END_VAR
VAR CONSTANT
	unWaitInterrupt						:UINT := 0;
	unDuringInterrupt						:UINT := 1;
	unAfterInterrupt						:UINT := 2;
	unChkFile							:UINT := 3;
	unNoInterrupt							:UINT := 4;
END_VAR

IF NOT bEnable
THEN
	bBusy := FALSE;
	bDone := FALSE;
	bError := FALSE;
	bEStop := FALSE;
	bFirstTime := FALSE;
	RETURN;
END_IF

IF NOT bFirstTime
THEN
	bBusy := FALSE;
	bDone := FALSE;
	bError := FALSE;
	bEStop := FALSE;
	unState := 0;
	unIncLog := 1;
	unIncDuringInterrupt := 1;
	unIncAfterInterrupt := 1;

	unLOG_INSTANCE_IDX  := GVL_Logger.unLOG_INSTANCE_IDX + 1;
	unInstanceIdx := unLOG_INSTANCE_IDX;

	unState := unWaitInterrupt;

	bFirstTime := TRUE;
END_IF


rtDeleteAll(CLK := bDeleteAll);

IF rtDeleteAll.Q
    AND (bDone OR bError)
THEN
	bBusy := FALSE;
	bDone := FALSE;
	bError := FALSE;
	bEStop := FALSE;
	unState := 0;
	unIncLog := 1;
	unIncDuringInterrupt := 1;
	unIncAfterInterrupt := 1;

	unState := unWaitInterrupt;
END_IF

rtInterrupt(CLK := bInterrupt);
IF rtInterrupt.Q
THEN
	unState := unWaitInterrupt;
END_IF;

udnCycleNo := udnCycleNo + 1;

CASE unState OF
	
	unWaitInterrupt:
		bBusy := FALSE;
		bDone := FALSE;
		bError := FALSE;

		fbLoggerFile.bExecute := FALSE;

		(* Shift down logger list by 1 *)
		A_ShiftDown();

		(* Write time stamp and value of variables before interrupt *)
		arstLoggerWaitInterrupt[1].udnCycleNo := udnCycleNo;
		arstLoggerWaitInterrupt[1].sTimeStamp := sDateTime;
		arstLoggerWaitInterrupt[1].arsLogVars := arsLogVars;

		IF bInterrupt
		THEN
			bBusy := TRUE;
			bDone := FALSE;

			bEStop := bLogOne;

			MEMSET(ADR(arstLoggerDuringInterrupt), 0, SIZEOF(arstLoggerDuringInterrupt));
			MEMSET(ADR(arstLoggerAfterInterrupt), 0, SIZEOF(arstLoggerAfterInterrupt));

			(* Log data *)
			IF unIncLog <= GVL_Logger.unLOG_MAX_NO
			THEN
				MEMCPY(ADR(arstLogger[unIncLog].arstLoggerWaitInterrupt), ADR(arstLoggerWaitInterrupt), SIZEOF(arstLoggerWaitInterrupt));
			ELSE
				unIncLog := 1;
				MEMCPY(ADR(arstLogger[unIncLog].arstLoggerWaitInterrupt), ADR(arstLoggerWaitInterrupt), SIZEOF(arstLoggerWaitInterrupt));
			END_IF

			(* Write time stamp and value of variables during interrupt *)
			unIncDuringInterrupt := 1;
			arstLoggerDuringInterrupt[unIncDuringInterrupt].udnCycleNo := udnCycleNo;
			arstLoggerDuringInterrupt[unIncDuringInterrupt].sTimeStamp := sDateTime;
			arstLoggerDuringInterrupt[unIncDuringInterrupt].arsLogVars := arsLogVars;
			unIncDuringInterrupt := unIncDuringInterrupt + 1;

			fbLoggerFile.sFileName := CONCAT(
										sDateTime,
										CONCAT(
											'_',
											UINT_TO_STRING(unInstanceIdx)
										)
									);

			unState := unDuringInterrupt;

		END_IF

	unDuringInterrupt:
		IF unIncDuringInterrupt <= GVL_Logger.unLOG_DURING_MAX_NO
		THEN
			(*  Write time stamp and value of variables during interrupt *)
			arstLoggerDuringInterrupt[unIncDuringInterrupt].udnCycleNo := udnCycleNo;
			arstLoggerDuringInterrupt[unIncDuringInterrupt].sTimeStamp := sDateTime;
			arstLoggerDuringInterrupt[unIncDuringInterrupt].arsLogVars := arsLogVars;
		
			unIncDuringInterrupt := unIncDuringInterrupt + 1;

		END_IF

		IF NOT bInterrupt
		THEN
			(* Log data *)
			MEMCPY(ADR(arstLogger[unIncLog].arstLoggerDuringInterrupt), ADR(arstLoggerDuringInterrupt), SIZEOF(arstLoggerDuringInterrupt));

			(* Write time stamp and value of variables after interrupt *)
			unIncAfterInterrupt := 1;
			arstLoggerAfterInterrupt[unIncAfterInterrupt].udnCycleNo := udnCycleNo;
			arstLoggerAfterInterrupt[unIncAfterInterrupt].sTimeStamp := sDateTime;
			arstLoggerAfterInterrupt[unIncAfterInterrupt].arsLogVars := arsLogVars;
			unIncAfterInterrupt := unIncAfterInterrupt + 1;

			unState := unAfterInterrupt;

		END_IF

	unAfterInterrupt:
		IF unIncAfterInterrupt <= GVL_Logger.unLOG_AFTER_MAX_NO
		THEN
			(* Write time stamp and value of variables after interrupt *)
			arstLoggerAfterInterrupt[unIncAfterInterrupt].udnCycleNo := udnCycleNo;
			arstLoggerAfterInterrupt[unIncAfterInterrupt].sTimeStamp := sDateTime;	
			arstLoggerAfterInterrupt[unIncAfterInterrupt].arsLogVars := arsLogVars;

			unIncAfterInterrupt := unIncAfterInterrupt + 1;
		ELSE
			(* Log data *)
			MEMCPY(ADR(arstLogger[unIncLog].arstLoggerAfterInterrupt), ADR(arstLoggerAfterInterrupt), SIZEOF(arstLoggerAfterInterrupt));

			fbLoggerFile.bExecute := TRUE;

			IF fbLoggerFile.bBusy
			THEN
				unState := unChkFile;

			ELSIF fbLoggerFile.bError
			THEN
				fbLoggerFile.bExecute := FALSE;
	
				bBusy := FALSE;
				bError := TRUE;
	
				unState := unNoInterrupt;

			END_IF
		END_IF

	unChkFile:
		IF NOT bEnableSaveInFile
		     OR fbLoggerFile.bDone
		THEN
			fbLoggerFile.bExecute := FALSE;

			bBusy := FALSE;
			bDone := TRUE;

			unState := unNoInterrupt;

		ELSIF  fbLoggerFile.bError
		THEN
			fbLoggerFile.bExecute := FALSE;

			bBusy := FALSE;
			bError := TRUE;

			unState := unNoInterrupt;

		END_IF

	unNoInterrupt:
		IF NOT bInterrupt
		    AND NOT bEStop
		THEN
			bBusy := FALSE;
			bDone := FALSE;
			bError := FALSE;

			unIncLog := unIncLog + 1;

			unState := unWaitInterrupt;
		END_IF

END_CASE


fbLoggerFile(
	bEnable := bEnableSaveInFile,
	sFilePath := sFilePath,
	sFileSuffix := sFileSuffix,
	arstLoggerWaitInterrupt := arstLoggerWaitInterrupt,
	arstLoggerDuringInterrupt := arstLoggerDuringInterrupt,
	arstLoggerAfterInterrupt := arstLoggerAfterInterrupt
 );

ACTION A_ShiftDown:

FOR nIdx := GVL_Logger.unLOG_BEFOR_MAX_NO - 1 TO 1 BY -1
DO
	arstLoggerWaitInterrupt[nIdx + 1] := arstLoggerWaitInterrupt[nIdx];
END_FOR
END_ACTION

END_FUNCTION_BLOCK

// ---- POUs/Tc3 Objects/Logic/F_DwordToBitReal_1.TcPOU
FUNCTION F_DwordToBitReal_1 : REAL
VAR_INPUT
	dwIn : DWORD;
END_VAR
VAR
	pt : POINTER TO REAL;
END_VAR

pt := ADR(dwIn);
F_DwordToBitReal := pt^;

END_FUNCTION

// ---- POUs/Tc3 Objects/Logic/F_RealToBitDword_1.TcPOU
FUNCTION F_RealToBitDword_1 : DWORD
VAR_INPUT
	rIn : REAL;
END_VAR
VAR
	pt : POINTER TO DWORD;
END_VAR

pt := ADR(rIn);
F_RealToBitDword := pt^;

END_FUNCTION

// ---- POUs/Tc3 Objects/Logic/F_ResetBitOfDWord_1.TcPOU
FUNCTION F_ResetBitOfDWord_1 : DWORD
VAR_INPUT
	dwInput			:DWORD;
	usnBitNr			:USINT;
END_VAR
VAR
END_VAR

F_ResetBitOfDWord := dwInput;
CASE usnBitNr OF
	0:
	F_ResetBitOfDWord.0 := FALSE;
	1:
	F_ResetBitOfDWord.1 := FALSE;
	2:
	F_ResetBitOfDWord.2 := FALSE;
	3:
	F_ResetBitOfDWord.3 := FALSE;
	4:
	F_ResetBitOfDWord.4 := FALSE;
	5:
	F_ResetBitOfDWord.5 := FALSE;
	6:
	F_ResetBitOfDWord.6 := FALSE;
	7:
	F_ResetBitOfDWord.7 := FALSE;
	8:
	F_ResetBitOfDWord.8 := FALSE;
	9:
	F_ResetBitOfDWord.9 := FALSE;
	10:
	F_ResetBitOfDWord.10 := FALSE;
	11:
	F_ResetBitOfDWord.11 := FALSE;
	12:
	F_ResetBitOfDWord.12 := FALSE;
	13:
	F_ResetBitOfDWord.13 := FALSE;
	14:
	F_ResetBitOfDWord.14 := FALSE;
	15:
	F_ResetBitOfDWord.15 := FALSE;
	16:
	F_ResetBitOfDWord.16 := FALSE;
	17:
	F_ResetBitOfDWord.17 := FALSE;
	18:
	F_ResetBitOfDWord.18 := FALSE;
	19:
	F_ResetBitOfDWord.19 := FALSE;
	20:
	F_ResetBitOfDWord.20 := FALSE;
	21:
	F_ResetBitOfDWord.21 := FALSE;
	22:
	F_ResetBitOfDWord.22 := FALSE;
	23:
	F_ResetBitOfDWord.23 := FALSE;
	24:
	F_ResetBitOfDWord.24 := FALSE;
	25:
	F_ResetBitOfDWord.25 := FALSE;
	26:
	F_ResetBitOfDWord.26 := FALSE;
	27:
	F_ResetBitOfDWord.27 := FALSE;
	28:
	F_ResetBitOfDWord.28 := FALSE;
	29:
	F_ResetBitOfDWord.29 := FALSE;
	30:
	F_ResetBitOfDWord.30 := FALSE;
	31:
	F_ResetBitOfDWord.31 := FALSE;
END_CASE

END_FUNCTION

// ---- POUs/Tc3 Objects/Logic/F_SetBitOfDWord_1.TcPOU
FUNCTION F_SetBitOfDWord_1 : DWORD
VAR_INPUT
	dwInput			:DWORD;
	usnBitNr			:USINT;
END_VAR
VAR
END_VAR

F_SetBitOfDWord := dwInput;
CASE usnBitNr OF
	0:
	F_SetBitOfDWord.0 := TRUE;
	1:
	F_SetBitOfDWord.1 := TRUE;
	2:
	F_SetBitOfDWord.2 := TRUE;
	3:
	F_SetBitOfDWord.3 := TRUE;
	4:
	F_SetBitOfDWord.4 := TRUE;
	5:
	F_SetBitOfDWord.5 := TRUE;
	6:
	F_SetBitOfDWord.6 := TRUE;
	7:
	F_SetBitOfDWord.7 := TRUE;
	8:
	F_SetBitOfDWord.8 := TRUE;
	9:
	F_SetBitOfDWord.9 := TRUE;
	10:
	F_SetBitOfDWord.10 := TRUE;
	11:
	F_SetBitOfDWord.11 := TRUE;
	12:
	F_SetBitOfDWord.12 := TRUE;
	13:
	F_SetBitOfDWord.13 := TRUE;
	14:
	F_SetBitOfDWord.14 := TRUE;
	15:
	F_SetBitOfDWord.15 := TRUE;
	16:
	F_SetBitOfDWord.16 := TRUE;
	17:
	F_SetBitOfDWord.17 := TRUE;
	18:
	F_SetBitOfDWord.18 := TRUE;
	19:
	F_SetBitOfDWord.19 := TRUE;
	20:
	F_SetBitOfDWord.20 := TRUE;
	21:
	F_SetBitOfDWord.21 := TRUE;
	22:
	F_SetBitOfDWord.22 := TRUE;
	23:
	F_SetBitOfDWord.23 := TRUE;
	24:
	F_SetBitOfDWord.24 := TRUE;
	25:
	F_SetBitOfDWord.25 := TRUE;
	26:
	F_SetBitOfDWord.26 := TRUE;
	27:
	F_SetBitOfDWord.27 := TRUE;
	28:
	F_SetBitOfDWord.28 := TRUE;
	29:
	F_SetBitOfDWord.29 := TRUE;
	30:
	F_SetBitOfDWord.30 := TRUE;
	31:
	F_SetBitOfDWord.31 := TRUE;
END_CASE

END_FUNCTION

// ---- POUs/Tc3 Objects/Logic/Oscat/CHECK_PARITY_1.TcPOU
FUNCTION CHECK_PARITY_1 : BOOL
(*
CHECK_PARITY checks an input byte IN and an associated paritybit P to
even parity. The output is TRUE if the number of bits in the byte IN have
the value TRUE together with the parity-bit results is an even number.
*)
VAR_INPUT
	in : DWORD;	(* input dword *)
	p : BOOL;	(* Parity-Bit *)
END_VAR


(*
version 1.3	18 feb 2008
programmer 	hugo
tested by	tobias

this function checks for an even partity for a dword and partity bit.

*)

CHECK_PARITY := NOT p;
WHILE in > 0 DO
	CHECK_PARITY := CHECK_PARITY XOR in.0 XOR in.1 XOR in.2 XOR in.3;
	in := SHR(in,4);
END_WHILE;

(* code before rev 1.2
WHILE in > 0 DO
	IF in.0 THEN cnt := cnt + 1; END_IF;
	in := SHR(in,1);
END_WHILE;
check_parity := even(cnt) XOR P;
*)


(* revision history

rev 1.0 HM  1.oct.2006

rev 1.1 hm	10.sep.2007
	changed algorithm to improove performance

rev 1.2	hm	8 dec 2007
	changed algorithm to improove performance

rev 1.3 hm	18. feb 2008
	changed algorithm to improove performance
*)

END_FUNCTION

// ---- POUs/Tc3 Objects/Mathematical/Delay/FB_Delay_1.TcPOU
FUNCTION_BLOCK FB_Delay_1
(*
Function block used to caculate delay

Constructor: 		Patryk Panylo
Company:		E. Riexinger GmbH
Date:			14.07.2014
Version:			1.00

Date:			Revision:		Who:				Comment
dd.mm.yyyy		x.xx			Initials			comment

*)
VAR_INPUT
	(* Enummerations *)

	(* Variables *)
	bEnable								:BOOL := TRUE;					(* Enable FB *)

	lrInSignal								:LREAL;							(* Input signal *)
	tDeadTime							:TIME := t#200ms;					(* Dead time *)
	tTaskCycle							:TIME := t#10ms; 					(* Cycle time *)

	(* References *)

	(* Interfaces *)

	(* Instances *)
END_VAR
VAR_OUTPUT
	(* Enummerations *)
	
	(* Variables *)
	lrOutSignal							:LREAL;							(* Output signal *)

	(* References *)

	(* Interfaces *)

	(* Instances *)
END_VAR
VAR
	(* Enummerations *)

	(* Variables *)
	bFirstTime							:BOOL;							(* First cycle *)

	lrTimeRatio							:LREAL;
	lrLastSignal							:LREAL;							(* Last signal *)

	(* References *)

	(* Interfaces *)

	(* Instances *)
	tpClock								:TP;

END_VAR

IF NOT bEnable
THEN
	lrOutSignal := lrInSignal;

	bFirstTime := FALSE;
	RETURN;
END_IF

IF NOT bFirstTime
THEN
	lrOutSignal := lrInSignal;

	tpClock(
		IN := FALSE,
		PT := tTaskCycle
	);

	bFirstTime := TRUE;
END_IF


tpClock();

IF NOT tpClock.Q
THEN
	tpClock(IN := FALSE);

	IF tDeadTime > t#0ms
	THEN
		lrTimeRatio := TIME_TO_LREAL(tTaskCycle) / TIME_TO_LREAL(tDeadTime);

		lrOutSignal := lrLastSignal + (lrInSignal - lrLastSignal) * lrTimeRatio;
	ELSE
		lrOutSignal := lrLastSignal;
	END_IF

	tpClock(IN := TRUE);
END_IF

lrLastSignal := lrOutSignal;

END_FUNCTION_BLOCK

// ---- POUs/Tc3 Objects/Mathematical/FB_Differential_1.TcPOU
FUNCTION_BLOCK FB_Differential_1
(*
Function block used to calculate differential

Constructor: 		Patryk Panylo
Company:		E. Riexinger GmbH
Date:			05.06.2014
Version:			1.00

Date:			Revision:		Who:				Comment
dd.mm.yyyy		x.xx			Initials			comment

*)
VAR_INPUT
	(* Enummerations *)
	
	(* Variables *)
	bEnable								:BOOL := TRUE;					(* Enable FB *)

	lrInSignal								:LREAL;							(* Input signal *)
	lrDifferentialValue						:LREAL := 1.0;						(* Differential value *)
	lrTaskCycle							:LREAL := 1.0; 					(* Cycle time *)

	(* References *)

	(* Interfaces *)

	(* Instances *)
END_VAR
VAR_OUTPUT
	(* Enummerations *)
	
	(* Variables *)
	lrOutSignal							:LREAL;							(* Output signal *)

	(* References *)

	(* Interfaces *)

	(* Instances *)
END_VAR
VAR
	(* Enummerations *)
	
	(* Variables *)
	bFirstTime							:BOOL;							(* First cycle *)

	lrLastSignal							:LREAL;							(* Last signal *)

	(* References *)

	(* Interfaces *)

	(* Instances *)


END_VAR

IF NOT bEnable
THEN
	lrOutSignal := lrInSignal;

	bFirstTime := FALSE;
	RETURN;
END_IF

IF NOT bFirstTime
THEN
	lrLastSignal := lrInSignal;
	bFirstTime := TRUE;
END_IF

IF lrTaskCycle > 0.0
THEN
	lrOutSignal := lrDifferentialValue * (lrInSignal - lrLastSignal) / lrTaskCycle;
ELSE
	lrOutSignal := 0.0;
END_IF
lrLastSignal := lrInSignal;

END_FUNCTION_BLOCK

// ---- POUs/Tc3 Objects/Mathematical/FB_Integral_1.TcPOU
FUNCTION_BLOCK FB_Integral_1
(*
Function block used to calculate integral

Constructor: 		Patryk Panylo
Company:		E. Riexinger GmbH
Date:			05.06.2014
Version:			1.00

Date:			Revision:		Who:				Comment
dd.mm.yyyy		x.xx			Initials			comment

*)
VAR_INPUT
	(* Enummerations *)

	(* Variables *)
	bEnable								:BOOL := TRUE;					(* Enable FB *)

	lrInSignal								:LREAL;							(* Input signal *)
	lrIntegralValue						:LREAL := 1.0;						(* Integration value in 1/sec *)
	lrTaskCycle							:LREAL := 1.0; 					(* Cycle time *)

	(* References *)

	(* Interfaces *)

	(* Instances *)
END_VAR
VAR_OUTPUT
END_VAR
VAR_IN_OUT
	(* Enummerations *)
	
	(* Variables *)
	lrOutSignal							:LREAL;							(* Output signal *)

	(* References *)

	(* Interfaces *)

	(* Instances *)
END_VAR
VAR
	(* Enummerations *)
	
	(* Variables *)
	bFirstTime							:BOOL;							(* First cycle *)

	lrLastSignal							:LREAL;							(* Last signal *)

	(* References *)

	(* Interfaces *)

	(* Instances *)


END_VAR

IF NOT bEnable
THEN
	bFirstTime := FALSE;
	RETURN;
END_IF

IF NOT bFirstTime
THEN
	lrLastSignal := lrInSignal;
	bFirstTime := TRUE;
END_IF

lrOutSignal := lrIntegralValue * lrTaskCycle * (lrInSignal + lrLastSignal) * 0.5 + lrOutSignal;
lrLastSignal := lrInSignal;

END_FUNCTION_BLOCK

// ---- POUs/Tc3 Objects/Mathematical/F_Exp10_1.TcPOU
FUNCTION F_Exp10_1 : REAL
VAR_INPUT
	X : REAL;
END_VAR


(*
version 1.0	 2 dec 2007
programmer 	hugo
tested by		tobias

this function calculates the exponent to the basis 10
exp10(3) = 1000

*)

F_Exp10 := EXP(X * 2.30258509299405);

END_FUNCTION

// ---- POUs/Tc3 Objects/Mathematical/F_FloorDN_1.TcPOU
FUNCTION F_FloorDN_1 : DINT
(*
Rounding down function which returns the biggest double integer.

Constructor: 		Patryk Panylo
Company:		E. Riexinger GmbH
Date:			20.01.2014
Version:			1.00

Date:			Revision:		Who:				Comment
dd.mm.yyyy		x.xx			Initials			comment

*)
VAR_INPUT
	rInValue						:REAL;
END_VAR
VAR
END_VAR


F_FloorDN := REAL_TO_DINT(rInValue);

IF DINT_TO_REAL(F_FloorDN) > rInValue
THEN
	F_FloorDN := F_FloorDN - 1;
END_IF

END_FUNCTION

// ---- POUs/Tc3 Objects/Mathematical/F_FracR_1.TcPOU
FUNCTION F_FracR_1 : REAL
(*
Function used to get fraction part of a real number.

Constructor: 		Patryk Panylo
Company:		E. Riexinger GmbH
Date:			17.07.2014
Version:			1.00

Date:			Revision:		Who:				Comment
dd.mm.yyyy		x.xx			Initials			comment

*)
VAR_INPUT
	(* Enummerations *)

	(* Variables *)
	rReal 						:REAL;			(* Input variable *)

	(* References *)

	(* Interfaces *)

	(* Instances *)

END_VAR
VAR
	(* Enummerations *)
	
	(* Variables *)
	rFloor						:REAL;

	(* References *)

	(* Interfaces *)

	(* Instances *)

END_VAR


rFloor := DINT_TO_REAL(F_FloorDN(ABS(rReal)));								(* Floor the value *)

IF rReal < 0
THEN
	F_FracR := rReal + rFloor ;								(* The fraction of the value *)

ELSE
	F_FracR := rReal - rFloor;								(* The fraction of the value *)

END_IF

END_FUNCTION

// ---- POUs/Tc3 Objects/Mathematical/F_GCD_1.TcPOU
FUNCTION F_GCD_1 : INT
(* Greatest common divisor *)
VAR_INPUT
	A : DINT;
	B : DINT;
END_VAR
VAR
	t: DINT;
END_VAR


(*
version 1.0	19. jan. 2011
programmer 	hugo
tested by	tobias

this function calculates the gretaest common divisor of two numbers A and B

*)

IF A = 0 THEN
	F_GCD := DINT_TO_INT(ABS(B));
ELSIF B = 0 THEN
	F_GCD := DINT_TO_INT(ABS(A));
ELSE
	A := ABS(A);
	B := ABS(B);
	F_GCD := 1;
	WHILE NOT(A.0 OR B.0) DO
		A := SHR(A,1);
		B := SHR(B,1);
		F_GCD := SHL(F_GCD,1);
	END_WHILE;
	WHILE A > 0 DO
		IF NOT(A.0) THEN A := SHR(A,1);
		ELSIF NOT(B.0) THEN B := SHR(B,1);
		ELSE
			t:= SHR(ABS(A-B),1);
			IF A < B THEN B := t; ELSE A := T; END_IF;
		END_IF;
	END_WHILE;
	F_GCD := F_GCD * DINT_TO_INT(B);
END_IF;


(* revision history
hm	19. jan. 2011	rev 1.0
	original version

*)

END_FUNCTION

// ---- POUs/Tc3 Objects/Mathematical/F_LRealRound_1.TcPOU
FUNCTION F_LRealRound_1 : LREAL
(*

The function used to round lreal value.

Constructor: 		Patryk Panylo
Company:		E. Riexinger GmbH
Date:			04.08.2015
Version:			1.00

Date:			Revision:		Who:				Comment
dd.mm.yyyy		x.xx			Initials			comment

*)
VAR_INPUT
	(* Input variables / Eingang Variablen *)
	lrReal							:LREAL; 						(*  Input variable *)
	usiPrecision						:USINT := 2; 					(* The number of digits after the decimal point depends on the requested precision *)
END_VAR
VAR
	(* Variables *)
	lrFraction							:LREAL;
END_VAR

(* Round real value with precision *)
lrFraction := FRAC(ABS(lrReal)) * EXPT(10, usiPrecision + 1); 							(* The fraction of the value *)

IF LMOD(lrFraction, 10) < 5
THEN
	lrFraction := lrFraction - LMOD(lrFraction, 10) ;										(* Round down *)
ELSE
	lrFraction := lrFraction + (10 - LMOD(lrFraction, 10));									(* Round up and check the integral increment *)
END_IF;

IF lrReal  < 0																		(* Check the digit of the value *)
THEN
	F_LRealRound	 := LTRUNC(lrReal) - (lrFraction / EXPT(10, usiPrecision + 1));
ELSE
	F_LRealRound	 := LTRUNC(lrReal) + (lrFraction / EXPT(10, usiPrecision + 1));
END_IF

END_FUNCTION

// ---- POUs/Tc3 Objects/Mathematical/F_ModDW_1.TcPOU
FUNCTION F_ModDW_1 : DWORD
(*
Modulo function for double word numbers (dividend mod divisor).

Constructor: 		Patryk Panylo
Company:		E. Riexinger GmbH
Date:			20.01.2014
Version:			1.00

Date:			Revision:		Who:				Comment
dd.mm.yyyy		x.xx			Initials			comment

*)
VAR_INPUT
	dwDividend						:DWORD;
	dwDivisor						:DWORD;
END_VAR
VAR
END_VAR


F_MODDW := dwDivisor;

IF dwDivisor <> 0 
THEN
	F_MODDW := dwDividend MOD dwDivisor;
END_IF;

END_FUNCTION

// ---- POUs/Tc3 Objects/Mathematical/F_ModR_1.TcPOU
FUNCTION F_ModR_1 : REAL
(*
Modulo function for real numbers (dividend mod divisor).

Constructor: 		Patryk Panylo
Company:		E. Riexinger GmbH
Date:			20.01.2014
Version:			1.00

Date:			Revision:		Who:				Comment
dd.mm.yyyy		x.xx			Initials			comment

*)
VAR_INPUT
	rDividend						:REAL;
	rDivisor							:REAL := 1.0;
END_VAR
VAR
END_VAR


F_ModR := rDivisor;

IF rDivisor <> 0.0 
THEN
	F_ModR := rDividend - DINT_TO_REAL(F_FloorDN(rDividend / rDivisor)) * rDivisor;
END_IF;

END_FUNCTION

// ---- POUs/Tc3 Objects/Mathematical/F_RoundR_1.TcPOU
FUNCTION F_RoundR_1 : REAL
(*
Function used to round real value with precision

Constructor: 		Patryk Panylo
Company:		E. Riexinger GmbH
Date:			17.07.2014
Version:			1.00

Date:			Revision:		Who:				Comment
dd.mm.yyyy		x.xx			Initials			comment

*)
VAR_INPUT
	(* Enummerations *)
	
	(* Variables *)
	rReal 						:REAL;			(* Input variable *)
	usnPrecision					:USINT := 2;		(* The number of digits after the decimal point depends on the requested precision *)

	(* References *)

	(* Interfaces *)

	(* Instances *)

END_VAR
VAR
	(* Enummerations *)
	
	(* Variables *)
	rFraction						:REAL;

	(* References *)

	(* Interfaces *)

	(* Instances *)

END_VAR


rFraction := F_FracR(ABS(rReal)) * EXPT(10, usnPrecision + 1); 								(* The fraction of the value *)

IF F_ModR(rFraction, 10) < 5
THEN
	rFraction := rFraction - F_ModR(rFraction, 10) ;											(* Round down *)
ELSE
	rFraction := rFraction + (10 - F_ModR(rFraction, 10));										(* Round up and check the integral increment *)
END_IF;

IF rReal  < 0																			(* Check the digit of the value *)
THEN
	F_RoundR := TRUNC(rReal) - (rFraction / EXPT(10, usnPrecision + 1));
ELSE
	F_RoundR := TRUNC(rReal) + (rFraction / EXPT(10, usnPrecision + 1));
END_IF

END_FUNCTION

// ---- POUs/Tc3 Objects/Mathematical/Hysteresis/FB_Hysteresis_1.TcPOU
FUNCTION_BLOCK FB_Hysteresis_1
(*
Function block used to generate hysteresis

Constructor: 		Patryk Panylo
Company:		E. Riexinger GmbH
Date:			15.07.2016
Version:			1.00

Date:			Revision:		Who:				Comment
dd.mm.yyyy		x.xx			Initials			comment

*)
VAR_INPUT
	(* Enummerations *)

	(* Variables *)
	bEnable							:BOOL := TRUE;					(* Enable FB *)

	lrInSignal							:LREAL;							(* Input signal *)
	lrGoDown						:REAL;
	lrGoUp							:REAL;

	(* References *)

	(* Interfaces *)

	(* Instances *)
END_VAR
VAR_OUTPUT
	(* Enummerations *)
	
	(* Variables *)
	lrOutSignal						:LREAL;						(* Output signal *)
	bLowLevel						:BOOL;						(* Low level detected *)
	bGoLevel						:BOOL;						(* Go level detected *)
	bHighLevel						:BOOL;						(* High level detected *)

	(* References *)

	(* Interfaces *)

	(* Instances *)
END_VAR
VAR
	(* Enummerations *)

	(* Variables *)
	bFirstTime							:BOOL;							(* First cycle *)

	lrLastSignal							:LREAL;							(* Last signal *)

	(* References *)

	(* Interfaces *)

	(* Instances *)

END_VAR

IF NOT bEnable
THEN
	lrOutSignal := lrInSignal;

	bFirstTime := FALSE;
	RETURN;
END_IF

IF NOT bFirstTime
THEN

	bFirstTime := TRUE;
END_IF

lrOutSignal:=SEL(lrInSignal - lrGoUp > lrLastSignal, lrOutSignal, lrInSignal - lrGoUp);
lrOutSignal:=SEL(lrInSignal + lrGoDown < lrLastSignal, lrOutSignal, lrInSignal + lrGoDown);

lrLastSignal := lrOutSignal;

END_FUNCTION_BLOCK

// ---- POUs/Tc3 Objects/Mathematical/Limits/FB_Limiter_1.TcPOU
FUNCTION_BLOCK FB_Limiter_1
(*
Function block used to limits input signal. 

Constructor: 		Patryk Panylo
Company:		E. Riexinger GmbH
Date:			21.07.2014
Version:			1.00

Date:			Revision:		Who:				Comment
dd.mm.yyyy		x.xx			Initials			comment

*)
VAR_INPUT
	(* Enummerations *)

	(* Variables *)
	bEnable								:BOOL := TRUE;					(* Enable FB *)

	lrInSignal								:LREAL;							(* Input signal *)
	lrLimitMin								:LREAL;							(* Limit minimum *)
	lrLimitMax							:LREAL;							(* Limit maximum *)

	(* References *)

	(* Interfaces *)

	(* Instances *)
END_VAR
VAR_OUTPUT
	(* Enummerations *)
	
	(* Variables *)
	lrOutSignal							:LREAL;							(* Output signal *)
	bLimitMin							:BOOL;							(* Minimum limit reached *)
	bLimitMax							:BOOL;							(* Maximum limit reached *)

	(* References *)

	(* Interfaces *)

	(* Instances *)
END_VAR
VAR
	(* Enummerations *)
	
	(* Variables *)
	bFirstTime							:BOOL;							(* First cycle *)

	(* References *)

	(* Interfaces *)

	(* Instances *)

END_VAR

IF NOT bEnable
THEN
	lrOutSignal := lrInSignal;

	bLimitMin := FALSE;							(* Minimum limit reached *)
	bLimitMax := FALSE;							(* Maximum limit reached *)

	bFirstTime := FALSE;
	RETURN;
END_IF

IF NOT bFirstTime
THEN

	bFirstTime := TRUE;
END_IF

lrOutSignal := lrInSignal;
bLimitMin := FALSE;							(* Minimum limit reached *)
bLimitMax := FALSE;							(* Maximum limit reached *)

IF lrInSignal <= lrLimitMin
THEN
	lrOutSignal  := lrLimitMin;
	bLimitMin := TRUE;

ELSIF lrInSignal >= lrLimitMax
THEN
	lrOutSignal := lrLimitMax;
	bLimitMax := TRUE;

END_IF

END_FUNCTION_BLOCK

// ---- POUs/Tc3 Objects/Mathematical/Limits/F_DeadZone_1.TcPOU
FUNCTION F_DeadZone_1 : REAL
(*
Function used to calculate dead zone.

Constructor: 		Patryk Panylo
Company:		E. Riexinger GmbH
Date:			03.06.2014
Version:			1.00

Date:			Revision:		Who:				Comment
dd.mm.yyyy		x.xx			Initials			comment

*)

VAR_INPUT
	(* Enummerations *)

	(* Variables *)
	lrInSignal								:LREAL;							(* Input signal *)
	lrDeadZone							:LREAL;							(* Dead zone *)

	(* References *)

	(* Interfaces *)

	(* Instances *)

END_VAR
VAR
	(* Enummerations *)

	(* Variables *)

	(* References *)

	(* Interfaces *)

	(* Instances *)

END_VAR


IF ABS(lrInSignal) > lrDeadZone
THEN
	F_DeadZone := lrInSignal;
ELSE
	F_DeadZone := 0.0;
END_IF;

END_FUNCTION

// ---- POUs/Tc3 Objects/Mathematical/Limits/F_WordToRange_1.TcPOU
FUNCTION F_WordToRange_1 : REAL
VAR_INPUT
	wWord 					:WORD;
	rLowLimit 				:REAL;
	rHighLimit 				:REAL;
END_VAR
VAR
END_VAR


F_WordToRange := (rHighLimit - rLowLimit) * WORD_TO_REAL(wWord) * 0.00001525902189669640 + rLowLimit;

END_FUNCTION

// ---- POUs/Tc3 Objects/Mathematical/Scaling/FB_ScalingOffset_1.TcPOU
FUNCTION_BLOCK FB_ScalingOffset_1
(*

The function block used to scaling input signal.

Constructor: 		Patryk Panylo
Company:		E. Riexinger GmbH
Date:			04.08.2015
Version:			1.00

Date:			Revision:		Who:				Comment
dd.mm.yyyy		x.xx			Initials			comment

*)
VAR_INPUT
	(* Input variables / Eingang Variablen *)
	bEnable							:BOOL;						(* Function block enable *)
	lrInput							:LREAL;						(* Input scaling proces value *)
	lrXLowLimit						:LREAL;						(* Upper limit of X range *)
	lrXUpperLimit						:LREAL; 						(*Upper limit of X range  *)
	lrYLowLimit						:LREAL; 						(* Low limit of Y range  *)
	lrYUpperLimit						:LREAL; 						(* Upper limit of Y range  *)
	usiPrecision						:USINT := 2; 					(* The number of digits after the decimal point depends on the requested precision *)
	lrOffset							:LREAL;						(* Offset of output *)
END_VAR
VAR_OUTPUT
	(* Output variables / Ausgang Variablen *)
	lrOutputRV						:LREAL;						(* Raw Value *)
	lrOutputPV						:LREAL;						(* Judgment Value  *)
END_VAR
VAR
	(* Instances / Instanzen *)
	fbScaling						:FB_Scaling;

	(* Enumerator  *)

	(* General flags / Allgemeine Variablen *)

END_VAR
VAR CONSTANT

END_VAR

IF NOT bEnable THEN
	fbScaling(
		bEnable := FALSE,
	);

	lrOutputRV := 0.0;					(* Raw Value *)
	lrOutputPV := 0.0;					(* Judgment Value *)
	RETURN;
END_IF

(* Scaling *)

fbScaling(
	bEnable := TRUE,
	lrInput := lrInput,
	lrXLowLimit := lrXLowLimit,
	lrXUpperLimit := lrXUpperLimit,
	lrYLowLimit := lrYLowLimit,
	lrYUpperLimit := lrYUpperLimit,
	usiPrecision := usiPrecision
);

lrOutputRV := fbScaling.lrOutputRV + lrOffset;
lrOutputPV := fbScaling.lrOutputPV + lrOffset;

END_FUNCTION_BLOCK

// ---- POUs/Tc3 Objects/Mathematical/Scaling/FB_Scaling_1.TcPOU
FUNCTION_BLOCK FB_Scaling_1
(*

The function block used to scaling input signal.

Constructor: 		Patryk Panylo
Company:		E. Riexinger GmbH
Date:			04.08.2015
Version:			1.00

Date:			Revision:		Who:				Comment
dd.mm.yyyy		x.xx			Initials			comment

*)
VAR_INPUT
	(* Input variables / Eingang Variablen *)
	bEnable							:BOOL;						(* Function block enable *)
	lrInput							:LREAL;						(* Input scaling proces value *)
	lrXLowLimit						:LREAL;						(* Upper limit of X range *)
	lrXUpperLimit						:LREAL; 						(*Upper limit of X range  *)
	lrYLowLimit						:LREAL; 						(* Low limit of Y range  *)
	lrYUpperLimit						:LREAL; 						(* Upper limit of Y range  *)
	usiPrecision						:USINT := 2; 					(* The number of digits after the decimal point depends on the requested precision *)
END_VAR
VAR_OUTPUT
	(* Output variables / Ausgang Variablen *)
	lrOutputRV						:LREAL;						(* Raw Value *)
	lrOutputPV						:LREAL;						(* Judgment Value  *)
	bLowLevel						:BOOL;						(* Low level detected *)
	bGoLevel						:BOOL;						(* Go level detected *)
	bHighLevel						:BOOL;						(* High level detected *)
END_VAR
VAR
	(* Instances / Instanzen *)

	(* Enumerator  *)

	(* General flags / Allgemeine Variablen *)
	lra								:LREAL;
	lrb								:LREAL;
END_VAR
VAR CONSTANT

END_VAR

IF NOT bEnable THEN
	lrOutputRV := 0.0;					(* Raw Value *)
	lrOutputPV := 0.0;					(* Judgment Value *)
	bLowLevel := FALSE;				(* Low level detected *)
	bGoLevel := FALSE;					(* Go level detected *)
	bHighLevel := FALSE;				(* High level detected *)
	RETURN;
END_IF

(* Scaling *)
IF lrInput > lrXUpperLimit															(* Check upper limit of X range *)
THEN
	lrOutputRV := lrYUpperLimit;
	bLowLevel := FALSE;
	bHighLevel := TRUE;
	bGoLevel := FALSE;
ELSIF lrInput <= lrXLowLimit														(* Check low limit of X range *)
THEN
	lrOutputRV := lrYLowLimit;
	bLowLevel := TRUE;
	bHighLevel := FALSE;
	bGoLevel := FALSE;
ELSE
	IF (((lrXUpperLimit - lrXLowLimit) < 0.01)											(* Check X range *)
	    AND ((lrXUpperLimit - lrXLowLimit) > -0.01))
	THEN
		lrOutputRV := lrYLowLimit;
		bLowLevel := TRUE;
		bHighLevel := FALSE;
		bGoLevel := FALSE;
	ELSE
		lra := (lrYUpperLimit - lrYLowLimit) / (lrXUpperLimit - lrXLowLimit);					(* Slope of a straight line, drawed by the range positions *)
		lrb := lrYUpperLimit - lra * lrXUpperLimit;
		lrOutputRV := lra * lrInput + lrb;
		bLowLevel := FALSE;
		bHighLevel := FALSE;
		bGoLevel := TRUE;
	END_IF;
END_IF

lrOutputPV := F_LRealRound(lrOutputRV, usiPrecision);

END_FUNCTION_BLOCK

// ---- POUs/Tc3 Objects/Measurements/Counter/FB_Counter_1.TcPOU
FUNCTION_BLOCK FB_Counter_1
VAR_INPUT
	(* Input variables / Eingang Variablen *)
	bEnable					:BOOL;						(* Enable FB signal *)
	bExecute				:BOOL;						(* Execute signal *)
	bReset					:BOOL;						(* Reset counter *)
END_VAR
VAR_OUTPUT
	(* Output variables / Ausgang Variablen *)
	bOverflow				:BOOL;						(* Overflow *)
	bAlarm					:BOOL;						(* Alarm signal *)
END_VAR
VAR_IN_OUT
	udnCounter				:UDINT;						(* Counter *)
END_VAR
VAR
	(* Enummerations *)

	(* Variables *)


	(* References *)

	(* Interfaces *)

	(* Instances *)
	rtCount					:R_TRIG;
	rtReset					:R_TRIG;

END_VAR

IF NOT bEnable
THEN

    RETURN;
END_IF;

rtReset(CLK := bReset);                    (* Reset rising edge *)

IF rtReset.Q                               		(* Count reset came *)
THEN
	udnCounter := 0;
END_IF;


rtCount(CLK := bExecute);                   		 (* Trigger rising edge *)

IF rtCount.Q                              		  		 (* Count trigger came *)
THEN
	IF udnCounter = 16#FFFFFFFF		 (* Detect counter overflow *)
	THEN
	    	bOverflow := TRUE;                  	 (* Counter overflow *)
	ELSE
	   	 bOverflow := FALSE;              	   	 (* Not counter overflow *)
	END_IF;
	
	udnCounter := udnCounter + 1;            	 (* Increment counter *)
END_IF;

END_FUNCTION_BLOCK

// ---- POUs/Tc3 Objects/Measurements/Counter/FB_DistanceCounter_1.TcPOU
FUNCTION_BLOCK FB_DistanceCounter_1
(*

Function block to read and write elapsed distance in/from file.
If sFileName or sFilePath  or sFileSuffix is empty then save function is diabled and generate error.

Constructor: 		Patryk Panylo
Company:		E. Riexinger GmbH
Date:			24.03.2014
Version:			1.00

Date:			Revision:		Who:				Comment
dd.mm.yyyy		x.xx			Initials			comment

*)

VAR_INPUT
	(* Variables *)
	bEnable							:BOOL;							(* Enable FB *)
	sAmsNetId 						:STRING := ''; 						(* Ams Net ID of file to read/write *)
	lrDistance						:LREAL; 							(* All over counter distance *)
	bCount							:BOOL; 							(* If true then count distance else save current distance *)
	bSave							:BOOL;							(* Save current distance counter *)
	bReset							:BOOL; 							(* Reset counter *)
	bDeleteAll						:BOOL; 							(* Delete all counters since beginning *)
	sFilePath						:STRING := 'C:\TwinCAT\Plc\';		(* File path *)
	sFileName						:STRING := 'default';				(* File name *)
	tSaveIntervall						:TIME := t#3m;						(* Intervall to save counter hours. If equal 0 then intervall is off *)
	tTimeout							:TIME := t#3s;						(* ADS timeout *)
END_VAR
VAR_OUTPUT
	(* Variables *)
	lrAllOverDistance					:LREAL; 							(* All over counter distance *)
	lrAfterResetDistance				:LREAL; 							(* Counter distance since last reset *)
	lrNoRetainDistance				:LREAL; 							(* No retain counter distance *)
	bError							:BOOL;							(* Program error *)
	udnErrNo						:UDINT;							(* Error number *)
END_VAR
VAR
	(* Enummerations *)
	etRWStep						:(eReadDistance, eChkRead, eWFWrite, eWriteDistance, eChkWrite, eError );

	(* Variables *)
	bFirstTime						:BOOL;
	stRetainDistance					:ST_DistanceCounter;
	stCacheRetainDistance			:ST_DistanceCounter;

	(* Instances *)
	ftCount							:F_TRIG;
	rtSave							:R_TRIG;
	rtReset							:R_TRIG;
	rtDeleteAll						:R_TRIG;

	fbFileHandler						:FB_FileHandlerBinary;				(* File handler *)
	tonWriteIntervall					:TON;							(* Timer for Save intervall control *)

END_VAR

IF NOT bEnable				(* Enable FB *)
THEN
	fbFileHandler(
		bEnable := FALSE,
		bExecute := FALSE,
		bFileRead := FALSE,
		bFileWrite := FALSE
	);

	bFirstTime := FALSE;
	bError := FALSE;			(* Program error *)
	udnErrNo := 0;				(* Error number *)

	RETURN;
END_IF


IF NOT bFirstTime
THEN
	(* Produce the file directory name *)
	fbFileHandler.sFilePath := sFilePath;
	fbFileHandler.sFileName := sFileName;
	fbFileHandler.sFileSuffix := 'dc';

	tonWriteIntervall(
		IN := FALSE,
		PT:= tSaveIntervall
	);

	etRWStep := eReadDistance;

	bFirstTime := TRUE;
	RETURN;
END_IF


(* Read / Write all over distance *)
CASE etRWStep OF

	eReadDistance:
		fbFileHandler.bExecute := TRUE;
		fbFileHandler.bFileRead := TRUE;
		fbFileHandler.bFileWrite := FALSE;

		IF fbFileHandler.bBusy
		THEN
			etRWStep := eChkRead;

		END_IF

	eChkRead:
		IF NOT fbFileHandler.bBusy
		THEN
			IF  fbFileHandler.bError
			THEN
				fbFileHandler.bExecute := FALSE;
				fbFileHandler.bFileRead := FALSE;
				fbFileHandler.bFileWrite := FALSE;

				stCacheRetainDistance.lrAllOverDistance := 0;
				stCacheRetainDistance.lrAfterResetDistance := 0;

				etRWStep := eWFWrite;				(* Next step *)

			ELSE
				fbFileHandler.bExecute := FALSE;
				fbFileHandler.bFileRead := FALSE;
				fbFileHandler.bFileWrite := FALSE;

				stCacheRetainDistance.lrAllOverDistance := stRetainDistance.lrAllOverDistance;
				stCacheRetainDistance.lrAfterResetDistance := stRetainDistance.lrAfterResetDistance;

				etRWStep := eWFWrite;				(* Next step *)

			END_IF
		END_IF

	eWFWrite:
		ftCount(
			CLK :=  bCount AND NOT bReset AND NOT bDeleteAll
		);

		rtSave(
			CLK := bSave AND NOT bReset AND NOT bDeleteAll
		);


		tonWriteIntervall(IN := tSaveIntervall > t#0s);

		IF ftCount.Q
		     OR rtSave.Q
		     OR tonWriteIntervall.Q
		THEN
			tonWriteIntervall(IN := FALSE);

			etRWStep := eWriteDistance;								(* Next step *)

		END_IF

	eWriteDistance:
		fbFileHandler.bExecute := TRUE;
		fbFileHandler.bFileRead := FALSE;
		fbFileHandler.bFileWrite := TRUE;

		IF fbFileHandler.bBusy
		THEN
			etRWStep := eChkWrite;								(* Next step *)

		END_IF

	eChkWrite:
		IF NOT fbFileHandler.bBusy
		THEN
			IF  fbFileHandler.bError
			THEN
				etRWStep := eError;								(* Next step *)

			ELSE
				fbFileHandler.bExecute := FALSE;
				fbFileHandler.bFileRead := FALSE;
				fbFileHandler.bFileWrite := FALSE;

				etRWStep := eWFWrite;							(* Next step *)

			END_IF
		END_IF

	eError:
		fbFileHandler.bExecute := FALSE;
		fbFileHandler.bFileRead := FALSE;
		fbFileHandler.bFileWrite := FALSE;

END_CASE


(* Counting distance *)
IF bCount
    AND NOT fbFileHandler.bFileRead
THEN
	lrNoRetainDistance := lrNoRetainDistance + lrDistance;
	stRetainDistance.lrAllOverDistance := stCacheRetainDistance.lrAllOverDistance + lrNoRetainDistance;
	stRetainDistance.lrAfterResetDistance := stCacheRetainDistance.lrAfterResetDistance + lrNoRetainDistance;
END_IF


(* Write / read  file *)
fbFileHandler(
	bEnable := TRUE,
	dwDataBuffer := ADR(stRetainDistance),
	udnDataBufLen := SIZEOF(stRetainDistance),
	tTimeout := tTimeout,
	bError => bError,
	udnErrNo => udnErrNo
);

rtReset(
	CLK := NOT bSave AND bReset
);
IF rtReset.Q
THEN
	stRetainDistance.lrAfterResetDistance := 0;
	lrNoRetainDistance := 0;
END_IF

rtDeleteAll(
	CLK := NOT bSave AND bDeleteAll
);
IF rtDeleteAll.Q
THEN
	stRetainDistance.lrAllOverDistance := 0;
	stRetainDistance.lrAfterResetDistance := 0;
	stCacheRetainDistance.lrAllOverDistance := 0;
	stCacheRetainDistance.lrAfterResetDistance := 0;
	lrNoRetainDistance := 0;
END_IF

(* Counter distance mapping *)
lrAllOverDistance := stRetainDistance.lrAllOverDistance;
lrAfterResetDistance := stRetainDistance.lrAfterResetDistance;

END_FUNCTION_BLOCK

// ---- POUs/Tc3 Objects/Measurements/Counter/FB_TimeHoursCounter_1.TcPOU
FUNCTION_BLOCK FB_TimeHoursCounter_1
(*

Function block to read and write elapsed time in/from file.
If sFileName or sFilePath  or sFileSuffix is empty then save function is diabled and generate error.

Constructor: 		Patryk Panylo
Company:		E. Riexinger GmbH
Date:			17.03.2014
Version:			1.00

Date:			Revision:		Who:				Comment
dd.mm.yyyy		x.xx			Initials			comment

*)

VAR_INPUT
	(* Variables *)
	bEnable							:BOOL;							(* Enable FB *)
	sAmsNetId 						:STRING := ''; 						(* Ams Net ID of file to read/write *)
	bCount							:BOOL; 							(* If true then count time else save current time *)
	bSave							:BOOL;							(* Save current hours counter *)
	bReset							:BOOL; 							(* Reset counter *)
	bDeleteAll						:BOOL; 							(* Delete all counters since beginning *)
	sFilePath						:STRING := 'C:\TwinCAT\Plc\';		(* File path *)
	sFileName						:STRING := 'default';				(* File name *)
	tSaveIntervall						:TIME := t#3m;						(* Intervall to save counter hours. If equal 0 then intervall is off *)
	tTimeout							:TIME := t#3s;						(* ADS timeout *)
END_VAR
VAR_OUTPUT
	(* Variables *)
	lrAllOverHours					:LREAL; 							(* All over counter hours *)
	lrAfterResetHours					:LREAL; 							(* Counter hours since last reset *)
	lrNoRetainHours					:LREAL; 							(* No retain counter hours *)
	bError							:BOOL;							(* Program error *)
	udnErrNo						:UDINT;							(* Error number *)
END_VAR
VAR
	(* Enummerations *)
	etRWStep						:(eReadHours, eChkRead, eWFWrite, eWriteHours, eChkWrite, eError );

	(* Variables *)
	bFirstTime						:BOOL;
	arlrCycleTimeAsHour				:ARRAY[0..2] OF LREAL;			(* Current cycle time as hours *)
	stRetainHours					:ST_TimeHoursCounter;

	(* Instances *)
	ftCount							:F_TRIG;
	rtSave							:R_TRIG;
	rtReset							:R_TRIG;
	rtDeleteAll						:R_TRIG;

	fbFileHandler						:FB_FileHandlerBinary;				(* File handler *)
	fbGetSystemTime					:GETSYSTEMTIME;				(* Detects System time *)
	tonWriteIntervall					:TON;							(* Timer for Save intervall control *)

END_VAR

IF NOT bEnable				(* Enable FB *)
THEN
	fbFileHandler(
		bEnable := FALSE,
		bExecute := FALSE,
		bFileRead := FALSE,
		bFileWrite := FALSE
	);

	bFirstTime := FALSE;
	bError := FALSE;			(* Program error *)
	udnErrNo := 0;				(* Error number *)

	RETURN;
END_IF


IF NOT bFirstTime
THEN
	(* Produce the file directory name *)
	fbFileHandler.sFilePath := sFilePath;
	fbFileHandler.sFileName := sFileName;
	fbFileHandler.sFileSuffix := 'thc';

	(* Get cycle time as hours *)
	A_GetCycleTime();

	tonWriteIntervall(
		IN := FALSE,
		PT:= tSaveIntervall
	);

	etRWStep := eReadHours;

	RETURN;
END_IF


(* Read / Write all over hours *)
CASE etRWStep OF

	eReadHours:
		fbFileHandler.bExecute := TRUE;
		fbFileHandler.bFileRead := TRUE;
		fbFileHandler.bFileWrite := FALSE;

		IF fbFileHandler.bBusy
		THEN
			etRWStep := eChkRead;

		END_IF

	eChkRead:
		IF NOT fbFileHandler.bBusy
		THEN
			IF  fbFileHandler.bError
			THEN
				fbFileHandler.bExecute := FALSE;
				fbFileHandler.bFileRead := FALSE;
				fbFileHandler.bFileWrite := FALSE;

				etRWStep := eWFWrite;				(* Next step *)

			ELSE
				fbFileHandler.bExecute := FALSE;
				fbFileHandler.bFileRead := FALSE;
				fbFileHandler.bFileWrite := FALSE;

				etRWStep := eWFWrite;				(* Next step *)

			END_IF
		END_IF

	eWFWrite:
		ftCount(
			CLK :=  bCount AND NOT bReset AND NOT bDeleteAll
		);

		rtSave(
			CLK := bSave AND NOT bReset AND NOT bDeleteAll
		);


		tonWriteIntervall(IN := tSaveIntervall > t#0s);

		IF ftCount.Q
		     OR rtSave.Q
		     OR tonWriteIntervall.Q
		THEN
			tonWriteIntervall(IN := FALSE);

			etRWStep := eWriteHours;								(* Next step *)

		END_IF

	eWriteHours:
		fbFileHandler.bExecute := TRUE;
		fbFileHandler.bFileRead := FALSE;
		fbFileHandler.bFileWrite := TRUE;

		IF fbFileHandler.bBusy
		THEN
			etRWStep := eChkWrite;								(* Next step *)

		END_IF

	eChkWrite:
		IF NOT fbFileHandler.bBusy
		THEN
			IF  fbFileHandler.bError
			THEN
				etRWStep := eError;								(* Next step *)

			ELSE
				fbFileHandler.bExecute := FALSE;
				fbFileHandler.bFileRead := FALSE;
				fbFileHandler.bFileWrite := FALSE;

				etRWStep := eWFWrite;							(* Next step *)

			END_IF
		END_IF

	eError:
		fbFileHandler.bExecute := FALSE;
		fbFileHandler.bFileRead := FALSE;
		fbFileHandler.bFileWrite := FALSE;

END_CASE


(* Counting hours *)
IF bCount
    AND NOT fbFileHandler.bFileRead
THEN
	stRetainHours.lrAllOverHours := stRetainHours.lrAllOverHours + arlrCycleTimeAsHour[0];
	stRetainHours.lrAfterResetHours := stRetainHours.lrAfterResetHours + arlrCycleTimeAsHour[0];
	lrNoRetainHours := lrNoRetainHours + arlrCycleTimeAsHour[0];
END_IF


(* Write / read  file *)
fbFileHandler(
	bEnable := TRUE,
	dwDataBuffer := ADR(stRetainHours),
	udnDataBufLen := SIZEOF(stRetainHours),
	tTimeout := tTimeout,
	bError => bError,
	udnErrNo => udnErrNo
);

rtReset(
	CLK := NOT bSave AND bReset
);
IF rtReset.Q
THEN
	stRetainHours.lrAfterResetHours := 0;
	//lrNoRetainHours := 0;
END_IF

rtDeleteAll(
	CLK := NOT bSave AND bDeleteAll
);
IF rtDeleteAll.Q
THEN
	stRetainHours.lrAllOverHours := 0;
	stRetainHours.lrAfterResetHours := 0;
	lrNoRetainHours := 0;
END_IF

(* Counter hours mapping *)
lrAllOverHours := stRetainHours.lrAllOverHours;
lrAfterResetHours := stRetainHours.lrAfterResetHours;

ACTION A_GetCycleTime:

(* Calculate system time *)
fbGetSystemTime();
arlrCycleTimeAsHour[0] := UINT64_TO_LREAL(IN := ULARGE_INTEGER(dwHighPart := fbGetSystemTime.timeHiDW, dwLowPart := fbGetSystemTime.timeLoDW))
									/ 10				(* Calculate into mycro seconds *)
									/ 1000			(* Calculate into millis econds *)
									/ 1000			(* Calculate into seconds *)
									/ 60				(* Calculate into minutes *)
									/ 60;				(* Calculate into hours *)


arlrCycleTimeAsHour[2] := arlrCycleTimeAsHour[1];
arlrCycleTimeAsHour[1] := arlrCycleTimeAsHour[0];

IF arlrCycleTimeAsHour[2] > 0
THEN
	arlrCycleTimeAsHour[0] := ABS(arlrCycleTimeAsHour[2] - arlrCycleTimeAsHour[1]);
	arlrCycleTimeAsHour[1] := 0;
	arlrCycleTimeAsHour[2] := 0;

	bFirstTime := TRUE;
END_IF
END_ACTION

END_FUNCTION_BLOCK

// ---- POUs/Tc3 Objects/Measurements/FB_MeanValue.TcPOU
FUNCTION_BLOCK FB_MeanValue
VAR_INPUT
	(* Input variables / Eingang Variablen *)
	bEnable					:BOOL;						(* Enable FB signal *)
	bReset					:BOOL;						(* Reset measurement *)
	bExecute				:BOOL;						(* Execute measurement *)
	bAbort					:BOOL;						(* Abort measurement *)
	lrSampleValue			:LREAL;						(* Sample measurement value *)
	lrSampleValueMin		:LREAL;						(* Sample measurement value minimum *)
	lrSampleValueMax		:LREAL;						(* Sample measurement value maximum *)
	udnSampleTime			:UDINT := 100;				(* Sample time [ms] *)
	udnSampleDeathStart		:UDINT;						(* Amount of death sample from start *)
	tMaxTime				:TIME := T#1092M;			(* Maximum time *)
END_VAR
VAR_OUTPUT
	(* Output variables / Ausgang Variablen *)
	lrMeanValue				:LREAL;						(* Mean measurement value *)
END_VAR
VAR_IN_OUT

END_VAR
VAR
	(* Enummerations *)

	(* Variables *)
	udnCounter				:UDINT;
	lrTotalValue			:LREAL;						(* Total measurement value *)
	bFirstTime				:BOOL;

	(* References *)

	(* Interfaces *)

	(* Instances *)
	fbCycleTime					:FB_Timer;
	
END_VAR

IF NOT bEnable
THEN
	lrMeanValue := lrSampleValue;
	bFirstTime := FALSE;
	RETURN;
END_IF;

IF NOT bFirstTime
THEN

	bFirstTime := TRUE;
END_IF;

(* Measuring time of cycle *)
fbCycleTime(
	bEnable := TRUE,
	bReset := bReset,
	bStartStop := bExecute,
	bStop := NOT bExecute OR bAbort,
	tMaxTime := tMaxTime
);

IF fbCycleTime.bTimeStarted 
THEN
	IF fbCycleTime.stActTime.dwMiliSec >= udnSampleTime * udnCounter
	THEN
		IF (lrSampleValue > lrSampleValueMin
			AND lrSampleValue < lrSampleValueMax)
			OR lrSampleValueMin = lrSampleValueMax
		THEN
			udnCounter := udnCounter + 1;
			
			IF udnCounter > udnSampleDeathStart
			THEN
				lrTotalValue := lrTotalValue + lrSampleValue;		
				lrMeanValue := lrTotalValue / UDINT_TO_LREAL(udnCounter - udnSampleDeathStart);
			END_IF
		END_IF		
	END_IF
ELSE
	lrTotalValue := 0;
	udnCounter := 0;
END_IF

END_FUNCTION_BLOCK

// ---- POUs/Tc3 Objects/Measurements/FB_TemperaturOK_1.TcPOU
FUNCTION_BLOCK FB_TemperaturOK_1
VAR_INPUT
	bEnable						:BOOL;			(* Enable FB signal *)
	bIn							:BOOL;			(* Temperature OK *)
	tTimeOutTempOK				:TIME := t#5s;		(* Temperature OK timeout *)
	tTimeOutTempNOK			:TIME := t#5s;		(* Temperature NOK timeout *)
END_VAR
VAR_OUTPUT
	bOut					:BOOL;			(* Temperature OK *)
	bError					:BOOL;			(* Error by temperature NOK *)
	udnErrorNo				:UDINT;
	udnMessageNo			:UDINT;
	sMsg					:STRING;
END_VAR
VAR
	bFirstTime			:BOOL;			(* First cycle *)
	tonDelayOK			:TON;			(* Temperatur delay ok *)
	tofWatchDog			:TOF;			(* Timer to off *)

END_VAR


IF NOT bFirstTime
THEN
	bError := FALSE;
	udnErrorNo := 0;
	udnMessageNo := 0;
	sMsg := '';
	tonDelayOK(
		IN := FALSE,
	          PT := tTimeOutTempOK
	);
	tofWatchDog(
		IN := FALSE,
	         PT := tTimeOutTempNOK
	);
	bFirstTime := TRUE;
END_IF;

(* Timer starts when came rising edge of signal *)
tonDelayOK(
	IN := bIn,
         PT := tTimeOutTempOK
);

tofWatchDog(
	IN := bIn,
         PT := tTimeOutTempNOK
);

IF tonDelayOK.Q
THEN
	bOut := TRUE;
    
ELSIF NOT tofWatchDog.Q
THEN
	bOut := FALSE;
    
END_IF;

END_FUNCTION_BLOCK

// ---- POUs/Tc3 Objects/Measurements/FB_Timer_1.TcPOU
FUNCTION_BLOCK FB_Timer_1
VAR_INPUT
	(* Input variables / Eingang Variablen *)
	bEnable					:BOOL;						(* Enable FB signal *)
	bReset					:BOOL;						(* Reset timer *)
	bStartStop				:BOOL;						(* Timer start stop *)
	bStop					:BOOL;						(* Timer stop *)
	tMaxTime				:TIME := t#1092m;				(* Maximum time *)
END_VAR
VAR_OUTPUT
	(* Output variables / Ausgang Variablen *)
	stRefTime				:ST_Time;						(* Reference time *)
	stActTime				:ST_Time;						(* Actuel time *)
	stRestTime				:ST_Time;						(* Rest time *)
END_VAR
VAR_IN_OUT

END_VAR
VAR
	(* Enummerations *)

	(* Variables *)
	stTime					:ST_Time;						(* Actuel time *)
	bTimeStarted			:BOOL;							(* Meassuare time started *)

	bFirstTime				:BOOL;

	(* References *)

	(* Interfaces *)

	(* Instances *)
	rtReset					:R_TRIG;
	rtStartStop				:R_TRIG;
	rtStop					:R_TRIG;

	tonMeassureTime			:TON;

END_VAR

IF NOT bEnable
THEN
	bTimeStarted := FALSE;
	rtStartStop(CLK := FALSE);
	tonMeassureTime(
		IN := FALSE,                   (* Reset timer *)
		PT := tMaxTime
	);

	bFirstTime := FALSE;
	RETURN;
END_IF;

IF NOT bFirstTime
THEN
	MEMSET(ADR(stActTime), 0, SIZEOF(stActTime));
	MEMSET(ADR(stRestTime), 0, SIZEOF(stRestTime));
	MEMSET(ADR(stTime), 0, SIZEOF(stTime));
	bFirstTime := TRUE;
END_IF;

IF bReset
THEN
	bTimeStarted := FALSE;
	tonMeassureTime(
		IN := FALSE,
	         PT := tMaxTime
	);
    
	MEMSET(ADR(stActTime), 0, SIZEOF(stActTime));
	MEMSET(ADR(stRestTime), 0, SIZEOF(stRestTime));
	MEMSET(ADR(stTime), 0, SIZEOF(stTime));
END_IF;


(* Rising edge start / stop *)
rtStartStop(CLK := bStartStop);

IF rtStartStop.Q                                   				 (* Startsignal trigger *)
THEN
	IF bTimeStarted                              			 (* Meassuare time started *)
	THEN
		bTimeStarted := TRUE;                      	 (* Time measure started *)
		tonMeassureTime(				 (* Stop (reset) timer *)
			IN := FALSE,
		         PT := tMaxTime
		);
		MEMSET(ADR(stTime), 0, SIZEOF(stTime));
	ELSE
		bTimeStarted := TRUE;                    	 (* Time measure started *)
		MEMSET(ADR(stTime), 0, SIZEOF(stTime));
	END_IF;
END_IF;

(* Rising edge stop*)
rtStop(CLK := bStop);

IF rtStop.Q                                        				 (* Stop timer *)
THEN
	bTimeStarted := FALSE;                        	 	 (* Time measure stoped *)
END_IF;

(* Start timer *)
tonMeassureTime(
	IN := bTimeStarted,
	PT := tMaxTime
);

(* Set outputs *)
stRefTime.dwSec := TIME_TO_DWORD(tonMeassureTime.PT) / 1000;

stRefTime.dwDeciSec := TIME_TO_DWORD(tonMeassureTime.PT) / 100;

stRefTime.dwCentiSec := TIME_TO_DWORD(tonMeassureTime.PT) / 10;

stRefTime.dwMiliSec := TIME_TO_DWORD(tonMeassureTime.PT) / 1;

IF bTimeStarted
THEN
	stActTime.dwSec := stTime.dwSec + TIME_TO_DWORD(tonMeassureTime.ET) / 1000;
	stRestTime.dwSec := TIME_TO_DWORD(tonMeassureTime.PT) / 1000 - stActTime.dwSec;
	
	stActTime.dwDeciSec := stTime.dwDeciSec + TIME_TO_DWORD(tonMeassureTime.ET) / 100;
	stRestTime.dwDeciSec := TIME_TO_DWORD(tonMeassureTime.PT) / 100 - stActTime.dwDeciSec;
	
	stActTime.dwCentiSec := stTime.dwCentiSec + TIME_TO_DWORD(tonMeassureTime.ET) / 10;
	stRestTime.dwCentiSec := TIME_TO_DWORD(tonMeassureTime.PT) / 10 - stActTime.dwCentiSec;

	stActTime.dwMiliSec := stTime.dwMiliSec + TIME_TO_DWORD(tonMeassureTime.ET) / 1;
	stRestTime.dwMiliSec := TIME_TO_DWORD(tonMeassureTime.PT) / 1 - stActTime.dwMiliSec;
END_IF;

IF tonMeassureTime.Q                                		(* Maximum time reached *)
THEN
	MEMSET(ADR(stTime), 0, SIZEOF(stTime));
	bTimeStarted := FALSE;                          		(* Time measure stoped *)
END_IF;

END_FUNCTION_BLOCK

// ---- POUs/Tc3 Objects/Measurements/Oscat/T_PLC_MS_1.TcPOU
FUNCTION T_PLC_MS_1 : DWORD
VAR CONSTANT
	debug			:BOOL := 0;
	N 				:INT := 0;
	offset 			:DWORD := 0;
END_VAR
VAR
	tx 				:TIME;
END_VAR

(*
version 1.2	16. nov 2008
programmer 	hugo
tested by	oscat

T_PLC_MS reads the internal PLC timer and return the time, it has the advantage to be able to set a debug mode 
and speed up the counter to test the plc timer overrun which occurs every 50 days respectively 25 days at siemens S7
this routine also allows to correct the behavior of s7 where the internal plc counter will not count all 32 bits.

*)

tx := TIME();
T_PLC_MS := TIME_TO_DWORD(Tx);
(* hier muss die korrektur für step7 stattfinden
plctime muss den vollen wertebereich von time ausnutzen:
wenn bei step7 time -24tage bis plus 24 tage ist dann muss der timer auch beim überlauf auf -24tage springen 
und auf keinen fall auf 0 !!!!
für siemens muss ein weiterer fb im main eingebunden werden der sicherstellt das alle 32 bits durchgezählt werden.
es kann nur ein fb sein den er muss sich das oberste (32te) bit merken.
oder etwa spring s7 bei überlauf auf -24 tage????? dann wäre keine korrektur nötig.
*)
IF debug
THEN
	T_PLC_MS := (SHL(T_PLC_MS,N) OR SHL(DWORD#1,N)-1) + OFFSET;
END_IF;

END_FUNCTION

// ---- POUs/Tc3 Objects/Measurements/RTC/FB_RTC_1.TcPOU
FUNCTION_BLOCK FB_RTC_1
VAR_INPUT
END_VAR
VAR_OUTPUT
	(* Variables *)
	bTimeValid							:BOOL;
	dtRTC        						:DT;
	dtRTCEX      						:DT;
	stDateTime							:ST_DateTime;
END_VAR
VAR
	(* Enummerations *)
	
	(* Variables *)
	bFirstTime							:BOOL;	
	bBusy								:BOOL;
	bError								:BOOL;
	udnErrorNo							:UDINT;			

	actSysTimeDate						:TIMESTRUCT;				(* Structure SysTimeDate *)
	
	bValidRTC      						:BOOL;	
	bValidRTCEX    						:BOOL;

	(* References *)

	(* Interfaces *)

	(* Instances *)

   	fbGetLocalTime  					:NT_GetTime;
	tonSyncTimer       					:TON;
	ftSyncTrigger     					:F_TRIG;

	rtFirstTime						:R_TRIG;

	fbRTC           						:RTC;
	fbRTCEX        						:RTC_EX;

	(* Information given by the RTC *)
	wYear								:WORD;
	wMonth								:WORD;
	wDay								:WORD;
	wHour								:WORD;
	wMinute								:WORD;
	wSecond							:WORD;
	wMilliseconds						:WORD;
	
	dtDatTimePunktHilfv :STRING;

END_VAR


IF NOT bFirstTime
THEN
	bFirstTime := TRUE;
	
END_IF


(* Get RTC *)
rtFirstTime(CLK := bFirstTime);

(* Time synchronization *)
tonSyncTimer(
	IN := NOT tonSyncTimer.Q,
	PT := T#100MS,
);

(* This function provides the time (seconds) which has passed since 01.01.1970 00:00:00 (RTC). *)
fbGetLocalTime(
	NETID := '',
	START := tonSyncTimer.Q
			 OR rtFirstTime.Q,
	TMOUT := T#5S,
	BUSY => bBusy,
	ERR => bError,
	ERRID => udnErrorNo
);

actSysTimeDate := fbGetLocalTime.TIMESTR;

(*This function converts the time given into format SysTimeDate.*)
ftSyncTrigger(CLK := bBusy AND NOT bError);

fbRTC(
	EN := ftSyncTrigger.Q, 
	PDT := SYSTEMTIME_TO_DT(actSysTimeDate), 
	Q => bValidRTC, 
	CDT => dtRTC 
);

fbRTCEX(
	EN := ftSyncTrigger.Q,
	PDT := SYSTEMTIME_TO_DT(actSysTimeDate),
	PMSEK := actSysTimeDate.wMilliseconds,
	Q => bValidRTCEX, 
	CDT => dtRTCEX 
);

(*The structure SysTimeDate contains detailed information on the system time, 
split up into a readable format, e.g.:*)

wYear := actSysTimeDate.wYear;
wMonth := actSysTimeDate.wMonth;
wDay := actSysTimeDate.wDay;
wHour := actSysTimeDate.wHour;
wMinute := actSysTimeDate.wMinute;
wSecond := actSysTimeDate.wSecond;
wMilliseconds := actSysTimeDate.wMilliseconds;

stDateTime.dtDateTime := dtRTC;
stDateTime.dtDateTimeEx := dtRTCEX;

stDateTime.sDate := CONCAT(WORD_TO_STRING(wYear),
		 CONCAT(SEL(LEN(WORD_TO_STRING(wMonth))=1 ,WORD_TO_STRING(wMonth),CONCAT('0',WORD_TO_STRING(wMonth))),
				SEL(LEN(WORD_TO_STRING(wDay))=1 ,WORD_TO_STRING(wDay),CONCAT('0',WORD_TO_STRING(wDay)))));

stDateTime.sTime := CONCAT(SEL(LEN(WORD_TO_STRING(wHour))=1 ,WORD_TO_STRING(wHour),CONCAT('0',WORD_TO_STRING(wHour))),
		 CONCAT(SEL(LEN(WORD_TO_STRING(wMinute))=1 ,WORD_TO_STRING(wMinute),CONCAT('0',WORD_TO_STRING(wMinute))),
				SEL(LEN(WORD_TO_STRING(wSecond))=1 ,WORD_TO_STRING(wSecond),CONCAT('0',WORD_TO_STRING(wSecond)))));

stDateTime.sTimeEx := CONCAT(stDateTime.sTime, SEL(LEN(WORD_TO_STRING(wMilliseconds))=1 , SEL(LEN(WORD_TO_STRING(wMilliseconds))=2 , WORD_TO_STRING(wMilliseconds), CONCAT('0',WORD_TO_STRING(wMilliseconds))), CONCAT('00',WORD_TO_STRING(wMilliseconds))));
				
stDateTime.sDateTime := CONCAT(stDateTime.sDate,CONCAT('_', stDateTime.sTime));

stDateTime.sDateTimeEx := CONCAT(stDateTime.sDate,CONCAT('_', stDateTime.sTimeEx));


dtDatTimePunktHilfv := DELETE(DT_TO_STRING(stDateTime.dtDateTime),4,0);
stDateTime.dtDateTimePunkt :=REPLACE(dtDatTimePunktHilfv,' ',1,11);

END_FUNCTION_BLOCK

// ---- POUs/Tc3 Objects/Safety/FB_AirPressure_1.TcPOU
FUNCTION_BLOCK FB_AirPressure_1
(*

The function block used to control air pressure.

Constructor: 		Patryk Panylo
Company:		E. Riexinger GmbH
Date:			23.04.2015
Version:			1.00

Date:			Revision:		Who:				Comment
dd.mm.yyyy		x.xx			Initials			comment

*)
VAR_INPUT
	(* Input variables / Eingang Variablen *)
	bEnable					:BOOL;						(* Enable FB signal *)
	bIn						:BOOL;						(* Input signal *)
	bNoEStop				:BOOL;						(* Emergency stop *)
	tAirOnDelay				:TIME := t#2s;					(* Delay air pressur on *)
	tTimeOut					:TIME := t#5s;					(* Timeout *)
END_VAR
VAR_OUTPUT
	(* Output variables / Ausgang Variablen *)
	bOut					:BOOL;						(* Air pressure ok *)
	bAirOn					:BOOL;						(* Air pressure on *)
	bError					:BOOL;						(* Error by no air pressure *)
	udnErrorNo				:UDINT;
	udnMessageNo			:UDINT;
	sMsg					:STRING;
END_VAR
VAR_IN_OUT

END_VAR
VAR
	(* Enummerations *)

	(* Variables *)
	bFirstTime				:BOOL;						(* First cycle *)

	(* References *)

	(* Interfaces *)

	(* Instances *)
	tonAirOnDelay			:TON;						(* Delay air pressur on *)
	tonWatchDog				:TON;						(* Timer to delay *)
END_VAR

IF NOT bEnable
THEN
	bOut := TRUE;
	bError := FALSE;
	udnErrorNo := 0;
	udnMessageNo := 0;
	sMsg := '';
	tonWatchDog(IN := FALSE,
	             		 PT := tTimeOut);
	bFirstTime := FALSE;
	RETURN;
END_IF;

IF NOT bFirstTime
THEN
	bError := FALSE;
	udnErrorNo := 0;
	udnMessageNo := 0;
	sMsg := '';
	tonWatchDog(IN := FALSE,
	             		 PT := tTimeOut);
	bFirstTime := TRUE;
END_IF;

tonAirOnDelay(
	IN := bNoEStop,
	PT := tAirOnDelay
);

bAirOn := tonAirOnDelay.Q;

(* Timer starts when came rising edge of signal *)
tonWatchDog(
	IN := bAirOn,
	PT := tTimeOut
);

bOut := bIn;
bError := NOT bOut
	        AND tonWatchDog.Q;

IF NOT bOut
     AND bAirOn
THEN
	IF tonWatchDog.Q                       		 (* Error if air pressure not present *)
	THEN
		udnErrorNo := 1;
		udnMessageNo := 0;
		sMsg := 'No pressured air';
	ELSE                                  				  (* Message if air pressure softstarting *)
		udnMessageNo := 1;
		sMsg := 'Air pressure building up';
	END_IF;
ELSE
	udnErrorNo := 0;
	udnMessageNo := 0;
	sMsg := '';
END_IF;

END_FUNCTION_BLOCK

// ---- POUs/Tc3 Objects/Safety/FB_LightCurtain_1.TcPOU
FUNCTION_BLOCK FB_LightCurtain_1
(*

The function block used to control light Curtain.

Constructor: 		Patryk Panylo
Company:		E. Riexinger GmbH
Date:			23.04.2015
Version:			1.00

Date:			Revision:		Who:				Comment
dd.mm.yyyy		x.xx			Initials			comment

*)
VAR_INPUT
	(* Input variables / Eingang Variablen *)
	bEnable					:BOOL;						(* Enable FB signal *)
	bIn						:BOOL;						(* Input signal *)
	bInConf					:BOOL;						(* Confirm *)
	tTimeOut					:TIME := t#1s;					(* Timeout *)
END_VAR
VAR_OUTPUT
	(* Output variables / Ausgang Variablen *)
	bOut					:BOOL;						(* Air pressure ok *)
	bOutConf					:BOOL;
	bError					:BOOL;						(* Error by no air pressure *)
	udnErrorNo				:UDINT;
	udnMessageNo			:UDINT;
	sMsg					:STRING;
END_VAR
VAR_IN_OUT

END_VAR
VAR
	(* Enummerations *)

	(* Variables *)
	bFirstTime				:BOOL;						(* First cycle *)

	(* References *)

	(* Interfaces *)

	(* Instances *)
	tonWatchDog				:TON;						(* Timer to delay *)
END_VAR

IF NOT bEnable
THEN
	bOut := TRUE;
	bError := FALSE;
	udnErrorNo := 0;
	udnMessageNo := 0;
	sMsg := '';
	tonWatchDog(IN := FALSE,
	             		 PT := tTimeOut);
	bFirstTime := FALSE;
	RETURN;
END_IF;

IF NOT bFirstTime
THEN
	bError := FALSE;
	udnErrorNo := 0;
	udnMessageNo := 0;
	sMsg := '';
	tonWatchDog(IN := FALSE,
				PT := tTimeOut);
	bFirstTime := TRUE;
END_IF;

(* Timer starts when came rising edge of signal *)
tonWatchDog(
	IN := bIn,
	PT := tTimeOut
);

bOut := tonWatchDog.Q;
bError := NOT bIn;

bOutConf := bInConf AND bError;

IF bError
THEN
	udnErrorNo := 1;
	sMsg := 'Light Curtain not ok';
    
ELSIF bOut
THEN
	udnErrorNo := 0;
	sMsg := 'Light curtain ok';
END_IF;

END_FUNCTION_BLOCK

// ---- POUs/Tc3 Objects/Safety/FB_NoEmergencyStop_1.TcPOU
FUNCTION_BLOCK FB_NoEmergencyStop_1
(*

The function block used to control emergency stop.

Constructor: 		Patryk Panylo
Company:		E. Riexinger GmbH
Date:			23.04.2015
Version:			1.00

Date:			Revision:		Who:				Comment
dd.mm.yyyy		x.xx			Initials			comment

*)
VAR_INPUT
	(* Input variables / Eingang Variablen *)
	bEnable					:BOOL;						(* Enable FB signal *)
	bIn						:BOOL;						(* Input signal *)
	bInConf					:BOOL;						(* Emergency stop *)
END_VAR
VAR_OUTPUT
	(* Output variables / Ausgang Variablen *)
	bOut					:BOOL;						(* Air pressure ok *)
	bOutConf					:BOOL;						(* Confirm output *)
	bError					:BOOL;						(* Error by no air pressure *)
	udnErrorNo				:UDINT;
	udnMessageNo			:UDINT;
	sMsg					:STRING;
END_VAR
VAR_IN_OUT

END_VAR
VAR
	(* Enummerations *)

	(* Variables *)
	bFirstTime				:BOOL;						(* First cycle *)

	(* References *)

	(* Interfaces *)

	(* Instances *)

END_VAR

IF NOT bEnable
THEN
	bOut := TRUE;
	bError := FALSE;
	udnErrorNo := 0;
	udnMessageNo := 0;
	sMsg := '';
	bFirstTime := FALSE;
	RETURN;
END_IF;

IF NOT bFirstTime
THEN
	bError := FALSE;
	udnErrorNo := 0;
	udnMessageNo := 0;
	sMsg := '';
	bFirstTime := TRUE;
END_IF;

bOut := bIn;
bError := NOT bOut;

IF bError
THEN
	udnErrorNo := 1;
	sMsg := 'Emergency stop';
ELSE
	udnErrorNo := 0;
	sMsg := 'No emergency stop';
END_IF;

bOutConf := bInConf AND NOT bIn;

END_FUNCTION_BLOCK

// ---- POUs/Tc3 Objects/Safety/FB_PowerSupply_1.TcPOU
FUNCTION_BLOCK FB_PowerSupply_1
(*

The function block used to control power supply.

Constructor: 		Patryk Panylo
Company:		E. Riexinger GmbH
Date:			23.04.2015
Version:			1.00

Date:			Revision:		Who:				Comment
dd.mm.yyyy		x.xx			Initials			comment

*)
VAR_INPUT
	(* Input variables / Eingang Variablen *)
	bEnable					:BOOL;						(* Enable FB signal *)
	bIn						:BOOL;						(* Input signal *)
	bNoEStop				:BOOL;						(* Emergency stop *)
	tPowerSupplyOn			:TIME := t#2s;					(* Timeout power supply on *)
	tPowerSupplyOff			:TIME := t#1s;					(* Timeout power supply off *)
END_VAR
VAR_OUTPUT
	(* Output variables / Ausgang Variablen *)
	bOut					:BOOL;						(* Power supply ok *)
	bError					:BOOL;						(* Error by no air pressure *)
	udnErrorNo				:UDINT;
	udnMessageNo			:UDINT;
	sMsg					:STRING;
END_VAR
VAR_IN_OUT

END_VAR
VAR
	(* Enummerations *)

	(* Variables *)
	bFirstTime				:BOOL;						(* First cycle *)

	(* References *)

	(* Interfaces *)

	(* Instances *)
	tonPowerSupplyOn		:TON;						(* Timer to delay *)
	tofPowerSupplyOff			:TOF;						(* Timer to delay *)
END_VAR

IF NOT bEnable
THEN
	bOut := TRUE;
	bError := FALSE;
	udnErrorNo := 0;
	udnMessageNo := 0;
	sMsg := '';
	tonPowerSupplyOn(IN := FALSE,
				            PT := tPowerSupplyOn);
	tofPowerSupplyOff(IN := FALSE,
	            			 PT := tPowerSupplyOff);
	bFirstTime := FALSE;
    RETURN;
END_IF;

IF NOT bFirstTime
THEN
	bError := FALSE;
	udnErrorNo := 0;
	udnMessageNo := 0;
	sMsg := '';
	tonPowerSupplyOn(IN := FALSE,
	          			  PT := tPowerSupplyOn);
	tofPowerSupplyOff(IN := FALSE,
	             			 PT := tPowerSupplyOff);
	bFirstTime := TRUE;
END_IF;

(* Timer starts when came rising edge of signal *)
tonPowerSupplyOn(
	IN := bIn AND bNoEStop,
         PT := tPowerSupplyOn
);

tofPowerSupplyOff(
	IN := tonPowerSupplyOn.Q AND bNoEStop,
         PT := tPowerSupplyOff
);

bOut := tofPowerSupplyOff.Q;
bError := NOT tofPowerSupplyOff.Q;

IF bError
THEN
	udnErrorNo := 1;
	udnMessageNo := 0;
	sMsg := 'No power supply';
ELSE
	udnErrorNo := 0;
	udnMessageNo := 0;
	sMsg := '';
END_IF;

END_FUNCTION_BLOCK

// ---- POUs/Tc3 Objects/Safety/FB_Temperature_1.TcPOU
FUNCTION_BLOCK FB_Temperature_1
(*

The function block used to control temperature.

Constructor: 		Patryk Panylo
Company:		E. Riexinger GmbH
Date:			23.04.2015
Version:			1.00

Date:			Revision:		Who:				Comment
dd.mm.yyyy		x.xx			Initials			comment

*)
VAR_INPUT
	(* Input variables / Eingang Variablen *)
	bEnable					:BOOL;						(* Enable FB signal *)
	bIn						:BOOL;						(* Input signal *)
	tTimeOut					:TIME := t#5s;					(* Timeout *)
END_VAR
VAR_OUTPUT
	(* Output variables / Ausgang Variablen *)
	bOut					:BOOL;						(* Air pressure ok *)
	bError					:BOOL;						(* Error by no air pressure *)
	bWarning				:BOOL;						(* Warning by no temperature *)
	udnErrorNo				:UDINT;
	udnMessageNo			:UDINT;
	sMsg					:STRING;
END_VAR
VAR_IN_OUT

END_VAR
VAR
	(* Enummerations *)

	(* Variables *)
	bFirstTime				:BOOL;						(* First cycle *)

	(* References *)

	(* Interfaces *)

	(* Instances *)
	tonWatchDog				:TON;						(* Timer to delay *)
END_VAR

IF NOT bEnable
THEN
	bOut := TRUE;
	bError := FALSE;
	udnErrorNo := 0;
	udnMessageNo := 0;
	sMsg := '';
	tonWatchDog(IN := FALSE,
	             		 PT := tTimeOut);
	bFirstTime := FALSE;
	RETURN;
END_IF;

IF NOT bFirstTime
THEN
	bError := FALSE;
	udnErrorNo := 0;
	udnMessageNo := 0;
	sMsg := '';
	tonWatchDog(IN := FALSE,
	             		 PT := tTimeOut);
	bFirstTime := TRUE;
END_IF;

(* Timer starts when came rising edge of signal *)
tonWatchDog(
	IN := NOT bIn,
	PT := tTimeOut
);

bOut := bIn;
bError := NOT bOut
	        AND tonWatchDog.Q;
bWarning := NOT bError
		      AND NOT bOut;

IF NOT bOut
THEN
	IF tonWatchDog.Q                       		 (* Error if air pressure not present *)
	THEN
		udnErrorNo := 1;
		udnMessageNo := 0;
		sMsg := 'Temperature not ok';
	END_IF;
ELSE
	udnErrorNo := 0;
	udnMessageNo := 0;
	sMsg := '';
END_IF;

END_FUNCTION_BLOCK

// ---- POUs/Tc3 Objects/Safety/Fieldbus/FB_Fieldbus_1.TcPOU
FUNCTION_BLOCK FB_Fieldbus_1
(*

The function block used to control fieldbus.

Constructor: 		Patryk Panylo
Company:		E. Riexinger GmbH
Date:			23.04.2015
Version:			1.00

Date:			Revision:		Who:				Comment
dd.mm.yyyy		x.xx			Initials			comment

*)
VAR_INPUT
	(* Input variables / Eingang Variablen *)
	bEnable					:BOOL;					(* Enable FB signal *)
	wFrmXWcState 			:WORD;					(* Link to task related ethercat frame state FrmXWcState *)
	nMasterDeviceId 			:UINT;
	nMasterSlaveCount		:UINT;
	nMasterSlaveCountCfg		:UINT;
	nMasterDevState			:UINT;
	arrMasterNetId			:T_AmsNetIdArr;
	tTimeOut					:TIME := t#5s;				(* Timeout for ADS commando *)
END_VAR
VAR_OUTPUT
	(* Output variables / Ausgang Variablen *)
	sMasterNetId				:T_AmsNetId ;			(* Fieldbus master ams net id*)
	bFieldbusOK				:BOOL;
	bFrameWcStateOK		:BOOL;
	bFrameWcStateError		:BOOL;
	bSlaveCountError			:BOOL;
	bMasterDevStateError		:BOOL;
	stMasterDevState			:ST_EcMasterDevState;
	bInit						:BOOL;
	bDone					:BOOL;					(* Program done *)
	bBusy					:BOOL;					(* Program busy  *)
	bError					:BOOL;					(* Program error  *)
	udnErrorNo				:UDINT;
	udnMessageNo			:UDINT;
	sMsg					:STRING;
END_VAR
VAR
	(* Enummerations *)

	(* Variables *)
	bFirstTime				:BOOL;
	wReqZeroMask			:WORD := 16#FFFF;		 (* Clear bit to ignore datagram error *)

	arstDiagSlaveInfo 			: ARRAY [0..3] OF ST_SlaveStateInfo;
	arstDiagSlaveInfoScanned	: ARRAY [0..3] OF ST_SlaveStateInfoScanned;

	(* References *)

	(* Interfaces *)

	(* Instances *)
	fbGetDeviceType			:IOF_GetDeviceType; 		(* Get the device type from the device ID *)
	fbEtherCATFrameDiag		:FB_EtherCATFrameDiag;
	fbEtherCATDiag			:FB_EtherCATDiag;
END_VAR

IF NOT bEnable
THEN
	fbGetDeviceType(START := FALSE);
	bFieldbusOK := FALSE;
	bFrameWcStateOK := FALSE;
	bFrameWcStateError := FALSE;
	bSlaveCountError := FALSE;
	bMasterDevStateError := FALSE;
	bInit := FALSE;
	bDone := FALSE;
	bBusy := FALSE;
	bError := FALSE;
	udnErrorNo := 0;
	udnMessageNo := 0;
	sMsg := '';
	RETURN;
END_IF;


IF NOT bFirstTime
THEN
	bFieldbusOK := FALSE;
	bFrameWcStateOK := FALSE;
	bFrameWcStateError := FALSE;
	bSlaveCountError := FALSE;
	bMasterDevStateError := FALSE;
	bInit := FALSE;
	bDone := FALSE;
	bBusy := FALSE;
	bError := FALSE;
	udnErrorNo := 0;
	udnMessageNo := 0;
	sMsg := '';
	bFirstTime := TRUE;
END_IF;

(* Get the device type from the device ID *)
fbGetDeviceType(
	NETID := '',
	DEVICEID := nMasterDeviceId,
	START := TRUE,
	TMOUT := tTimeOut
);

(* Get the device type from the device ID *)
IF NOT fbGetDeviceType.BUSY 										(* No error *)
     AND NOT fbGetDeviceType.ERR
THEN

	CASE fbGetDeviceType.IODeviceType
	OF
		48: (* IODEVICETYPE_FC7500 	:= 48,  Beckhoff-SERCOS-PCI *)
			bInit := TRUE;
			bDone := FALSE;
			bBusy := FALSE;
			bError := FALSE;
			udnErrorNo := 0;											(* Error number *)
			(*bInitReady := unMasterState = 16#E005; 						(* Actual Phase is 4 *)
			bBreak := unMasterState = 16#E008;							(* Interrupt / Broke *)*)

		94: (* IODEVICETYPE_EtherCAT := 94,  Beckhoff-EtherCAT-PCI *)
			sMasterNetId := F_CreateAmsNetId(nIds := arrMasterNetId);
			bInit := sMasterNetID <> '' AND sMasterNetID <> '0.0.0.0.0.0';

			fbEtherCATFrameDiag(
				wFrmXWcState := wFrmXWcState,
				wReqZeroMask := wReqZeroMask,
				bFrameWcStateOK => bFrameWcStateOK
			);


			fbEtherCATDiag(
				sNetID := '',
				sMasterNetID	 := sMasterNetId,
				nMasterDevID := nMasterDeviceId,
				nSlaveCount := nMasterSlaveCount,
				nSlaveCountCfg := nMasterSlaveCountCfg,
				nMasterDevState := nMasterDevState,
				bAllFrameWcStatesOK	:= bFrameWcStateOK,
				tTimeout := tTimeOut,
				arstDiagSlaveInfo := arstDiagSlaveInfo,
				arstDiagSlaveInfoScanned	:= arstDiagSlaveInfoScanned,
				bEtherCATOK => bFieldbusOK,
				bFrameWcStateError	=> bFrameWcStateError,
				bSlaveCountError	=> bSlaveCountError,
				bMasterDevStateError=> bMasterDevStateError,
				stMasterDevState	=> stMasterDevState,
				bDone => bDone,
				bBusy => bBusy,
				bError => bError,
				iErrorID => udnErrorNo
			);

	ELSE (* IDLE *)
		bInit := FALSE;
		bDone := FALSE;
		bBusy := FALSE;
		bError := TRUE;
		udnErrorNo := 1;																			(* Error number *)
		sMsg := CONCAT('Unidentified fieldbus:', DINT_TO_STRING(fbGetDeviceType.IODeviceType));		(* Description error *)
	END_CASE;

ELSIF NOT fbGetDeviceType.BUSY
	    AND fbGetDeviceType.ERR
THEN
	bInit := FALSE;
	bDone := FALSE;
	bBusy := FALSE;
	bError := TRUE;
	udnErrorNo := 2;																				(* Error number *)
	sMsg := CONCAT('Fehler beim Lesen über ADS: ', UDINT_TO_STRING(fbGetDeviceType.ERRID));		(* Description error *)
	fbGetDeviceType(START := FALSE);
END_IF;

END_FUNCTION_BLOCK

// ---- POUs/Tc3 Objects/Signals/Force Input/FB_ForceBit_1.TcPOU
FUNCTION_BLOCK FB_ForceBit_1
(*

Forcing the input bit through pointer.
IO variables in VAR_CONFIG are generated automatically by TwinCAT - read only
Matching variable must be with  %I* declarated.

Constructor: 		Patryk Panylo
Company:		E. Riexinger GmbH
Date:			28.10.2013
Version:			1.00

Date:			Revision:		Who:				Comment
dd.mm.yyyy		x.xx			Initials			comment

*)
VAR_INPUT
	bEnable						:BOOL; 							(* Enable FB *)
	dwBitAddr					:DWORD;						(* The address of input argument in a DWORD: BITADR(Input) where e.g Input = %IX0.1 *)
	bForceInState				:BOOL;							(* Force input state *)
	tDelayOn					:TIME;							(* Delay signal on *)
	tDelayOff					:TIME;							(* Delay signal off *)
END_VAR
VAR_OUTPUT
END_VAR
VAR
	pByteAddr					:POINTER TO BYTE;
	byCurrentInState				:BYTE;							(* Current input state *)
	byBitMask					:BYTE;

	tonDelayOn					:TON;
	tonDelayOff					:TOF;

END_VAR

IF NOT bEnable
THEN
	RETURN;
END_IF

(* Delay on signal *)
tonDelayOn(
	IN := bForceInState,
	PT := tDelayOn
);

(* Delay off signal *)
tonDelayOff(
	IN := tonDelayOn.Q,
	PT := tDelayOff
);

pByteAddr := ADR(%IB0) + (dwBitAddr / 8);
byCurrentInState := pByteAddr^;

byBitMask := SHL(BYTE#1, (dwBitAddr AND 2#00000111));

IF tonDelayOff.Q
THEN
	pByteAddr^ := byCurrentInState OR byBitMask;
ELSE
	pByteAddr^ := byCurrentInState AND NOT byBitMask;
END_IF

END_FUNCTION_BLOCK

// ---- POUs/Tc3 Objects/Signals/Force Input/FB_ForceByte_1.TcPOU
FUNCTION_BLOCK FB_ForceByte_1
(*

Forcing the input bit through pointer.
IO variables in VAR_CONFIG are generated automatically by TwinCAT - read only
Matching variable must be with  %I* declarated.

Constructor: 		Patryk Panylo
Company:		E. Riexinger GmbH
Date:			28.10.2013
Version:			1.00

Date:			Revision:		Who:				Comment
dd.mm.yyyy		x.xx			Initials			comment

*)
VAR_INPUT
	bEnable						:BOOL; 							(* Enable FB *)
	pByteAddr					:POINTER TO BYTE;				(* The address of input argument in a DWORD: ADR(Input) where e.g Input = %IB *)
	bForceInState				:BOOL;							(* Force input state *)
	tDelayOn					:TIME;							(* Delay signal on *)
	tDelayOff						:TIME;							(* Delay signal off *)
END_VAR
VAR_OUTPUT
END_VAR
VAR
	byCurrentInState				:BYTE;							(* Current input state *)
	byBitMask					:BYTE;

	tonDelayOn					:TON;
	tonDelayOff					:TOF;

END_VAR

IF NOT bEnable
THEN
	RETURN;
END_IF

(* Delay on signal *)
tonDelayOn(
	IN := bForceInState,
	PT := tDelayOn
);

(* Delay off signal *)
tonDelayOff(
	IN := tonDelayOn.Q,
	PT := tDelayOff
);

byCurrentInState := pByteAddr^;

byBitMask := 2#00000001;

IF tonDelayOff.Q
THEN
	pByteAddr^ := byCurrentInState OR byBitMask;
ELSE
	pByteAddr^ := byCurrentInState AND NOT byBitMask;
END_IF

END_FUNCTION_BLOCK

// ---- POUs/Tc3 Objects/Signals/Force Input/FB_ForceInput.TcPOU
FUNCTION_BLOCK FB_ForceInput
(*

Forcing the input bit through pointer.

Constructor: 		Patryk Panylo
Company:		E. Riexinger GmbH
Date:			04.04.2020
Version:			1.00

Date:			Revision:		Who:				Comment
dd.mm.yyyy		x.xx			Initials			comment

*)
VAR_INPUT
	bEnable						:BOOL; 							(* Enable FB *)
	pInputAddr					:POINTER TO BOOL;				(* The address of input argument *)
	bForceInState				:BOOL;							(* Force input state *)
	tDelayOn					:TIME;							(* Delay signal on *)
	tDelayOff					:TIME;							(* Delay signal off *)
END_VAR
VAR_OUTPUT
END_VAR
VAR
	pByteAddr					:POINTER TO BYTE;
	byCurrentInState				:BYTE;							(* Current input state *)
	byBitMask					:BYTE;

	tonDelayOn					:TON;
	tonDelayOff					:TOF;

END_VAR

IF NOT bEnable
THEN
	RETURN;
END_IF

(* Delay on signal *)
tonDelayOn(
	IN := bForceInState,
	PT := tDelayOn
);

(* Delay off signal *)
tonDelayOff(
	IN := tonDelayOn.Q,
	PT := tDelayOff
);

IF tonDelayOff.Q
THEN
	pInputAddr^ := TRUE;
ELSE
	pInputAddr^ := FALSE;
END_IF

END_FUNCTION_BLOCK

// ---- POUs/Tc3 Objects/Signals/Generators/FB_Blinker_1.TcPOU
FUNCTION_BLOCK FB_Blinker_1
(*

Frequency division

Constructor: 		Patryk Panylo
Company:		E. Riexinger GmbH
Date:			14.11.2012
Version:			1.00

Date:			Revision:		Who:				Comment
dd.mm.yyyy		x.xx			Initials			comment

*)

VAR_INPUT
	tPeriod				:TIME := T#250MS;				(* Blink period *)
	bReset				:BOOL;							(* Reset *)
END_VAR
VAR_OUTPUT
	stBlinker				:ST_Blinker;
END_VAR
VAR
	byInc				:BYTE;
	rtTriger				:R_TRIG;
	ton1					:TON;
	ton2					:TON;
END_VAR

IF bReset
THEN
	byInc := 0;

	ton1(IN := FALSE);
	ton2(IN := FALSE);

	stBlinker.Q0 := 0;
	stBlinker.Q1 := 0;
	stBlinker.Q2 := 0;
	stBlinker.Q3 := 0;
	stBlinker.Q4 := 0;
	stBlinker.Q5 := 0;
	stBlinker.Q6 := 0;
	stBlinker.Q7 := 0;
	
	RETURN;	
END_IF

ton1(IN := NOT ton2.Q, PT:= tPeriod/2);
ton2(IN := ton1.Q, PT := tPeriod/2);

rtTriger(CLK := ton1.Q);
IF rtTriger.Q THEN
	byInc := byInc + 1;
END_IF;

stBlinker.Q0 := byInc.0;
stBlinker.Q1 := byInc.1;
stBlinker.Q2 := byInc.2;
stBlinker.Q3 := byInc.3;
stBlinker.Q4 := byInc.4;
stBlinker.Q5 := byInc.5;
stBlinker.Q6 := byInc.6;
stBlinker.Q7 := byInc.7;

END_FUNCTION_BLOCK

// ---- POUs/Tc3 Objects/Signals/Handling/FB_SignalHandlingDelay_1.TcPOU
FUNCTION_BLOCK FB_SignalHandlingDelay_1
VAR_INPUT
	(* Input variables / Eingang Variablen *)
	bEnable					:BOOL;						(* Enable FB signal *)
	bIn						:BOOL;						(* Input signal *)
	tDelay					:TIME := t#0s;					(* Delay *)
END_VAR
VAR_OUTPUT
	(* Output variables / Ausgang Variablen *)
	bOut					:BOOL;						(* Delayed signal *)
END_VAR
VAR
	(* Enummerations *)

	(* Variables *)
	bFirstTime				:BOOL;						(* First cycle *)

	(* References *)

	(* Interfaces *)

	(* Instances *)
	tonDelay					:TON;						(* Timer to delay *)
END_VAR

IF NOT bEnable
THEN
	tonDelay(IN := FALSE,
	          	PT := tDelay);
	bOut := bIn;
    RETURN;
END_IF;

tonDelay(				(* Dealy input signal *)
	IN := bIn,
	PT := tDelay
);

bOut := tonDelay.Q;		(* Set output *)

END_FUNCTION_BLOCK

// ---- POUs/Tc3 Objects/Signals/Handling/FB_SignalHandlingEdge_1.TcPOU
FUNCTION_BLOCK FB_SignalHandlingEdge_1
VAR_INPUT
	(* Input variables / Eingang Variablen *)
	bEnable					:BOOL;						(* Enable FB signal *)
	bIn						:BOOL;						(* Input signal *)
	tDelay					:TIME := t#0s;					(* Delay *)
END_VAR
VAR_OUTPUT
	(* Output variables / Ausgang Variablen *)
	bOut					:BOOL;						(* Delayed signal *)
	bRisingEdge				:BOOL;						(* Rising edge *)
	bFallingEdge				:BOOL;						(* Falling edge *)
	bRisingEdgeDelay		:BOOL;						(* Rising edge delay *)
END_VAR
VAR
	(* Enummerations *)

	(* Variables *)


	(* References *)

	(* Interfaces *)

	(* Instances *)
	rtREdge					:R_TRIG;						(* Timer to delay *)
	rtREdgeDelay			:R_TRIG;						(* Timer to delay *)
	ftFEdge					:F_TRIG;						(* Timer to delay *)
	fbSignalHandlingDelay		:FB_SignalHandlingDelay;
END_VAR

IF NOT bEnable
THEN
	fbSignalHandlingDelay(
		bEnable := FALSE,
		bIn := bIn,
		bOut => bOut
	);

	rtREdge(CLK := FALSE);		(* Check rising edge *)
	ftFEdge(CLK := FALSE);		(* Check rising edge *)
	bRisingEdge := FALSE;
	bFallingEdge := FALSE;

	rtREdgeDelay(CLK := FALSE);		(* Check rising edge *)
	bRisingEdgeDelay := FALSE;
    RETURN;
END_IF;

fbSignalHandlingDelay(
	bEnable := TRUE,
	bIn := bIn,
	tDelay := tDelay,
	bOut => bOut
);

rtREdge(CLK := bIn);            			 (* Check rising edge *)
bRisingEdge := rtREdge.Q;

rtREdgeDelay(CLK := bOut);            			 (* Check rising edge *)
bRisingEdgeDelay := rtREdgeDelay.Q;

ftFEdge(CLK := bIn);            			 (* Check rising edge *)
bFallingEdge := ftFEdge.Q;

END_FUNCTION_BLOCK

// ---- POUs/Tc3 Objects/Signals/Handling/F_SignalHandling_1.TcPOU
FUNCTION F_SignalHandling_1 : BOOL
VAR_INPUT
	(* Input variables / Eingang Variablen *)
	bEnable					:BOOL;						(* Enable FB signal *)
	bIn						:BOOL;						(* Input signal *)
END_VAR
VAR
END_VAR

IF NOT bEnable
THEN
	F_SignalHandling := FALSE;
    	RETURN;
END_IF;

F_SignalHandling := bIn;                     (* Set output *)

END_FUNCTION

// ---- POUs/Tc3 Objects/Signals/Ramp Generators/FB_RampDirector_1.TcPOU
FUNCTION_BLOCK FB_RampDirector_1
(*

Frequency division

Constructor: 		Patryk Panylo
Company:		E. Riexinger GmbH
Date:			14.11.2012
Version:			1.00

Date:			Revision:		Who:				Comment
dd.mm.yyyy		x.xx			Initials			comment

*)

VAR_INPUT
	bEnable						:BOOL;						(* Function block enable *)
	bExecute					:BOOL;						(* Execut the function block *)
	bDirection					:BOOL;						(* Rising = 1, Falling = 0 *)
	bSet						:BOOL;						(* Set output to 65535 *)
	bReset						:BOOL;						(* Reset output to 0 *)
	tRiseTime					:TIME;						(* Rise time of ramp *)
	tFallTime					:TIME;						(* Fall time of ramp *)
	rHighLimit					:REAL;						(* High limit of ramp *)
	rLowLimit						:REAL;						(* Low limit of ramp *)
	rNoLimit						:REAL;						(* No limit value active if rise and fall time no active *)
END_VAR
VAR_OUTPUT
	wRVOut						:WORD;						(* Ramp value, 100% = 65535 *)
	rPVOut						:REAL;						(* Judgment Value *)
	nPVOut						:INT;						(* Judgment Value *)
	bLowLevel					:BOOL;						(* Low level reached *)
	bHighLevel					:BOOL;						(* High level reached *)
	bDone						:BOOL;						(* Program done *)
	bBusy 						:BOOL;						(* Program busy *)
	bError 						:BOOL;						(* Program error *)
END_VAR
VAR
	fbRampGen					:FB_RMP_W;					(* Ramp generator *)

	rCacheLowLimit				:REAL;
	rCacheHighLimit				:REAL;

	rtExecute						:R_TRIG;
	etRampGenerator				:ET_RampGenerator;
END_VAR


IF NOT bEnable
THEN
	bDone := FALSE;                                     (* Program done *)
	bBusy := FALSE;                                     (* Program not busy *)
	bError := FALSE;                                    (* Program not error *)
	
	rtExecute(CLK := FALSE);

	fbRampGen(
		bEnable := FALSE,
		bReset := bReset,
		bSet := bSet,
		wRVOut => wRVOut
	);

	RETURN;
END_IF;

rtExecute(CLK := bExecute);

IF rtExecute.Q
THEN
	fbRampGen(
		bEnable := FALSE,
		bDirection := bDirection,
		bSet := FALSE,
		bReset := FALSE,
		tRampTime := T#0ms
	);
	
	etRampGenerator := ET_RampGenerator_eWaitExecute;						(* Next step *)

END_IF

(* Reset ramp *)
IF (tFallTime = t#0s
    AND tRiseTime <> t#0s
    AND bExecute
    AND NOT bDirection)
    OR bReset
THEN
	fbRampGen.bReset := TRUE;
	wRVOut := fbRampGen.wRVOut;
ELSE
	fbRampGen.bReset := FALSE;
END_IF;

(* Set ramp *)
IF (tRiseTime = t#0s
    AND tFallTime <> t#0s
    AND bExecute
    AND bDirection)
    OR bSet
THEN
	fbRampGen.bSet := TRUE;
ELSE
	fbRampGen.bSet := FALSE;
END_IF;

(* Call ramp generator *)
fbRampGen(
	bDirection := bDirection,
	tRampTime := SEL(bDirection, tFallTime, tRiseTime),
	bLowLevel => bLowLevel,
	bHighLevel => bHighLevel
);

IF fbRampGen.bReset
    OR fbRampGen.bSet
THEN
	wRVOut := fbRampGen.wRVOut;
END_IF;

CASE etRampGenerator OF
        
	ET_RampGenerator_eWaitExecute:
		bDone := FALSE;                                     (* Program done *)
		bBusy := FALSE;                                     (* Program not  busy *)
		bError := FALSE;                                    (* Program not error *)

		fbRampGen.bEnable := FALSE;
		
		IF rtExecute.Q
		THEN
			bDone := FALSE;                                     (* Program done *)
			bBusy := TRUE;                                 	 	(* Program not busy *)

			IF tRiseTime = t#0s
    			     AND tFallTime = t#0s
			THEN
				fbRampGen.bEnable := FALSE;

				rCacheLowLimit := rNoLimit;
				rCacheHighLimit := rNoLimit;

				etRampGenerator := ET_RampGenerator_eDone;         (* Next step *)
			ELSE
				fbRampGen.bEnable := TRUE;

				rCacheLowLimit := rLowLimit;
				rCacheHighLimit := rHighLimit;

				etRampGenerator := ET_RampGenerator_eRunning;           (* Next step *)
			END_IF
		END_IF

	ET_RampGenerator_eRunning:
		IF fbRampGen.bBusy
		THEN
			wRVOut := fbRampGen.wRVOut;
		
			etRampGenerator := ET_RampGenerator_eWaiting;           (* Next step *)
		END_IF
        
	ET_RampGenerator_eWaiting:
		IF fbRampGen.bBusy
		THEN
			wRVOut := fbRampGen.wRVOut;
		ELSE
			fbRampGen.bEnable := FALSE;
		
			etRampGenerator := ET_RampGenerator_eDone;         (* Next step *)
		END_IF		

	ET_RampGenerator_eDone:
		bDone := TRUE;                                      (* Program done *)
		bBusy := FALSE;                                     (* Program not busy *)
		
		etRampGenerator := ET_RampGenerator_eNotExecute;            (* Next step *)
        
	ET_RampGenerator_eError:
		bDone := FALSE;                                     (* Program done *)
		bBusy := FALSE;                                     (* Program not busy *)
		bError := TRUE;                                     (* Program error *)
		
		etRampGenerator := ET_RampGenerator_eNotExecute;            (* Next step *)
        
	ET_RampGenerator_eNotExecute:
	IF NOT bExecute
	THEN
		bDone := FALSE;                                     (* Program done *)
		bBusy := FALSE;                                     (* Program not busy *)
		bError := FALSE;                                    (* Program not error *)

		wRVOut := fbRampGen.wRVOut;
	
		etRampGenerator := ET_RampGenerator_eWaitExecute;               (* Next step *)

	END_IF;
END_CASE;

rPVOut := F_WordToRange(
			wWord := wRVOut,
			rLowLimit := rCacheLowLimit,
			rHighLimit := rCacheHighLimit
		);

nPVOut := REAL_TO_INT(rPVOut);

END_FUNCTION_BLOCK

// ---- POUs/Tc3 Objects/Signals/Watchdog/FB_SignalWatchdogLimit.TcPOU
FUNCTION_BLOCK FB_SignalWatchdogLimit
VAR_INPUT
	bEnable					:BOOL;			(* Enable FB signal *)
	bIn						:BOOL;			(* Input *)
	tTimeOutHigh				:TIME := t#5s;		(* Input high timeout *)
	tTimeOutLow				:TIME := t#5s;		(* Input low timeout *)
END_VAR
VAR_OUTPUT
	bOut					:BOOL;			(* Output *)
	bError					:BOOL;			(* Error *)
	udnErrorNo				:UDINT;
	udnMessageNo			:UDINT;
	sMsg					:STRING;
END_VAR
VAR
	bFirstTime				:BOOL;			(* First cycle *)
	tonDelay					:TON;			(* Delay *)
	tofWatchDog				:TOF;			(* Timer to off *)

END_VAR


IF NOT bFirstTime
THEN
	bError := FALSE;
	udnErrorNo := 0;
	udnMessageNo := 0;
	sMsg := '';
	tonDelay(
		IN := FALSE,
	          PT := tTimeOutHigh
	);
	tofWatchDog(
		IN := FALSE,
	         PT := tTimeOutLow
	);
	bFirstTime := TRUE;
END_IF;

(* Timer starts when came rising edge of signal *)
tonDelay(
	IN := bIn,
         PT := tTimeOutHigh
);

tofWatchDog(
	IN := bIn,
         PT := tTimeOutLow
);

IF tonDelay.Q
THEN
	bOut := TRUE;
    
ELSIF NOT tofWatchDog.Q
THEN
	bOut := FALSE;
    
END_IF;

END_FUNCTION_BLOCK

// ---- POUs/Tc3 Objects/Signals/Watchdog/FB_SignalWatchdog_1.TcPOU
FUNCTION_BLOCK FB_SignalWatchdog_1
VAR_INPUT
	(* Input variables / Eingang Variablen *)
	bEnable					:BOOL;						(* Enable FB signal *)
	bIn						:BOOL;						(* Input signal *)
	tWatchdog				:TIME := t#0s;					(* Watchdog time *)
END_VAR
VAR_OUTPUT
	(* Output variables / Ausgang Variablen *)
	bOut					:BOOL;						(* Output signal *)
	bAlarm					:BOOL;						(* Alarm signal *)
END_VAR
VAR
	(* Enummerations *)

	(* Variables *)


	(* References *)

	(* Interfaces *)

	(* Instances *)
	tofWatchdog				:TOF;

END_VAR

IF NOT bEnable
THEN
	bOut := FALSE;
	bAlarm := FALSE;                       (* Alarm active *)
	
	tofWatchdog(
		IN := tofWatchdog.ET > t#0ms,
	         PT := t#0ms
	);
	
	tofWatchdog(IN := FALSE,
	             PT := t#0ms);

	RETURN;
END_IF;

tofWatchdog(					 (* Dealy input signal *)
	IN := bIn,
	PT := tWatchdog
);

bOut := tofWatchdog.Q;

bAlarm := NOT tofWatchdog.Q;                       (* Set alarm *)

END_FUNCTION_BLOCK

// ---- POUs/Tc3 Objects/String/F_CheckStringIsReal_1.TcPOU
FUNCTION F_CheckStringIsReal_1 : BOOL (* TRUE if STR does not contain capital letters *)
VAR_INPUT
	str : T_MaxString;
END_VAR
VAR
	L : INT;
	pt : POINTER TO BYTE;
	pt2 : POINTER TO BYTE;
	pos: INT;
	pos2: INT;
END_VAR

pt := ADR(str);
pt2 := ADR(str);
L := LEN(str);

FOR pos := 1 TO L DO

	IF pt^ = 43 (* + *)
	     AND (pos <> 1)
	THEN
		F_CheckStringIsReal := FALSE;
		RETURN;

	ELSIF pt^ = 44 (* , *)
	THEN
		IF (pos = 1 (*OR pos = L*))
		THEN
			F_CheckStringIsReal := FALSE;
			RETURN;
		ELSE
			FOR pos2 := 1 TO L DO
				IF pos <> pos2
				THEN
					IF pt2^ = 44 OR pt2^ = 46
					THEN
						F_CheckStringIsReal := FALSE;
						RETURN;
					END_IF
				END_IF
				pt2 := pt2 + 1;
			END_FOR
		END_IF;
	ELSIF pt^ = 45 (* - *)
	     AND (pos <> 1)
	THEN
		F_CheckStringIsReal := FALSE;
		RETURN;
	ELSIF pt^ = 46 (* . *)
	THEN
		IF (pos = 1 (*OR pos = L*))
		THEN
			F_CheckStringIsReal := FALSE;
			RETURN;
		ELSE
			FOR pos2 := 1 TO L DO
				IF pos <> pos2
				THEN
					IF pt2^ = 44 OR pt2^ = 46
					THEN
						F_CheckStringIsReal := FALSE;
						RETURN;
					END_IF
				END_IF
				pt2 := pt2 + 1;
			END_FOR
		END_IF;
	ELSIF NOT (pt^ > 47 AND pt^ < 58)	(* 0 .. 9 *)
	     	    AND pt^ <> 43 (* + *)
	    	    AND pt^ <> 44 (* , *)
	             AND pt^ <> 45 (* - *)
	     	    AND pt^ <> 46 (* . *)
	THEN
		F_CheckStringIsReal := FALSE;
		RETURN;
	END_IF;

    	pt := pt + 1;
END_FOR;
F_CheckStringIsReal := L > 0;

END_FUNCTION

// ---- POUs/Tc3 Objects/String/F_CheckSyntaxReal.TcPOU
FUNCTION F_CheckSyntaxReal : BOOL (* TRUE if STR does not contain capital letters *)
VAR_INPUT
	str 		:T_MaxString;
	flag 		:T_MaxString;
	sep 		:T_MaxString := '=';
	rsufix		:POINTER TO REAL; 					
END_VAR
VAR
	L			:INT;
	prefix1		:T_MaxString;
	prefix2		:T_MaxString;
	ssufix		:T_MaxString;
END_VAR


prefix1 := CONCAT(flag, sep);
L := LEN(prefix1);
prefix2 := MID(str, L, 1);

F_CheckSyntaxReal := FALSE;

IF LEN(str) > L
THEN
	ssufix := DELETE(str, L, 1);
	IF prefix1 = prefix2
	THEN
		IF F_CheckStringIsReal(ssufix)
		THEN
			F_CheckSyntaxReal := TRUE; 
			rsufix^ := STRING_TO_REAL(ssufix);
		END_IF
	END_IF;
END_IF

END_FUNCTION

// ---- POUs/Tc3 Objects/String/F_CheckSyntaxString.TcPOU
FUNCTION F_CheckSyntaxString : BOOL (* TRUE if STR does not contain capital letters *)
VAR_INPUT
	str 		:T_MaxString;
	flag 		:T_MaxString;
	sep 		:T_MaxString := '=';
	sufix		:POINTER TO STRING; 					
END_VAR
VAR
	L			:INT;
	prefix1		:T_MaxString;
	prefix2		:T_MaxString;
	
END_VAR


prefix1 := CONCAT(flag, sep);
L := LEN(prefix1);
prefix2 := MID(str, L, 1);

F_CheckSyntaxString := FALSE;

IF LEN(str) > L
THEN
	sufix^ := DELETE(str, L, 1);
	IF prefix1 = prefix2
	THEN
		F_CheckSyntaxString := TRUE;
	END_IF;
END_IF

END_FUNCTION

// ---- POUs/Tc3 Objects/String/F_RealToStrf_1.TcPOU
FUNCTION F_RealToStrf_1 : STRING(20)
VAR_INPUT
	IN : REAL;
	N : INT;
	D : STRING(1);
END_VAR
VAR
	O: REAL;
	i: INT;
END_VAR

(*
version 1.8	2. jan 2012
programmer 	hugo
tested by	oscat

Real_to_strf converts a Real to a fixed length String.
the string will be filles with zeroes to achieve the fixed length N after the decimal separator.
the input parameter specifies the decimal separator to be used in the output string.

*)

(* LIMIT N to 0 .. 7 *)
N := LIMIT(0,N,7);
(* round the input to N digits and convert to string *)
O := ABS(in) * F_Exp10(N);
F_RealToStrf := DINT_TO_STRING(REAL_TO_DINT(O));
(* add zeroes in front to make sure sting is at least 8 digits long *)
FOR i := LEN(F_RealToStrf) TO N DO F_RealToStrf := CONCAT('0', F_RealToStrf); END_FOR;
(* add a dot if n > 0 *)
IF n > 0 THEN F_RealToStrf := INSERT(F_RealToStrf, D, LEN(F_RealToStrf) - N); END_IF;
(* add a minus sign if in is negative *)
IF in < 0 THEN F_RealToStrf := CONCAT('-', F_RealToStrf); END_IF;

END_FUNCTION

// ---- POUs/Tc3 Objects/Traceability/FB_TraceCycle.TcPOU
FUNCTION_BLOCK FB_TraceCycle
(*

This function block is used to traceability of data.

Constructor: 		Patryk Panylo
Company:		E. Riexinger GmbH
Date:			02.09.2016
Version:			1.00

Date:			Revision:		Who:				Comment
21.02.2018		0.01			PPA						Additional logger for samples

*)
VAR_INPUT
	(* Input variables / Eingang Variablen *)
	bEnable						:BOOL;					(* Enable FB *)
	sFilePath					:STRING := 'C:\Riex\Traceability\NewData\';	(* Path to file e.g. 'c:\', \Hard Disk\ *)
	sFileName					:STRING := 'default';	(* Name of file *)
	bExecute					:BOOL;					(* Execute write data *)
	bAbort						:BOOL;					(* Abort write data *)
	bReset						:BOOL;					(* Reset write data *)			
	udnSampleTime				:UDINT := 100;			(* Sample time [ms] *)
	tMaxTime					:TIME := T#0S;			(* Maximal write time *)
	arsNameRecords				:ARRAY[0..GVL_Trace.MAX_TRACE_ROWS, 0..GVL_Trace.MAX_TRACE_COLUMNS] OF STRING(GVL_Trace.MAX_TRACE_FIELD_LENGTH);
	arsValueRecords				:ARRAY[0..GVL_Trace.MAX_TRACE_ROWS, 0..GVL_Trace.MAX_TRACE_COLUMNS] OF STRING(GVL_Trace.MAX_TRACE_FIELD_LENGTH);
	tTimeout					:TIME := T#1S;			(* States the time before the function is cancelled *)
END_VAR
VAR_OUTPUT
	(* Output variables / Ausgang Variablen *)
	bBusy						:BOOL;					(* Program busy *)
	bDone						:BOOL;					(* Program done *)
	bError						:BOOL;					(* Program error *)
	udnErrNo					:UDINT;					(* Error number *)
END_VAR
VAR_IN_OUT
	fbFileHandler				:FB_FileCSVHandler;				(* Traceability *)
END_VAR
VAR
	(* Enummerations *)
	etTraceState				:ET_TRACE_State := ET_TRACE_State_eWaitExecute;
	
	(* Variables *)
	udnWriteCounter				:UDINT;
	
	udnRowCounter				:UDINT;
	udnColumnCounter			:UDINT;

	bFirstTime					:BOOL;					(* First PLC cycle *)

	(* References *)

	(* Interfaces *)

	(* Instances *)
	rtExecute					:R_TRIG;
	fbCycleTime					:FB_Timer;
END_VAR

IF NOT bEnable				(* Enable FB *)
THEN
	bFirstTime := FALSE;		(* First PLC cycle *)
	bBusy := FALSE;			(* Program busy *)
	bDone := FALSE;			(* Program done *)
	bError := FALSE;			(* Program error *)
	udnErrNo := 0;				(* Error number *)
	RETURN;
END_IF

IF NOT bFirstTime
THEN

	bFirstTime := TRUE;
END_IF

IF bReset
   AND bError
THEN
	bBusy := FALSE;
	bDone := FALSE;
	bError := FALSE;
	
	fbCycleTime(bReset := TRUE);
	
	etTraceState := ET_TRACE_State_eWaitExecute;
END_IF

(* Measuring time of cycle *)
fbCycleTime(
	bEnable := TRUE,
	bReset := FALSE,
	bStartStop := bExecute,
	bStop := NOT bExecute OR bAbort,
	tMaxTime := tMaxTime
);

rtExecute(CLK := bExecute);

CASE etTraceState
OF
	ET_TRACE_State_eWaitExecute:
		IF rtExecute.Q
		   AND NOT fbFileHandler.bBusy
		THEN	
			bBusy := TRUE;
			bDone := FALSE;
			bError := FALSE;
			udnErrNo := 0;

			fbFileHandler.bExecute := FALSE;
			fbFileHandler.sFilePath := sFilePath;
			fbFileHandler.sFileName := sFileName; 
			
			udnWriteCounter := 0;
			udnRowCounter := 0;
			udnColumnCounter := 0;
			
			FOR udnRowCounter := 0 TO GVL_Trace.MAX_TRACE_ROWS
			DO 
				FOR udnColumnCounter := 0 TO GVL_Trace.MAX_TRACE_COLUMNS
				DO 
					fbFileHandler.arsWriteRecords[udnRowCounter, udnColumnCounter] := arsNameRecords[udnRowCounter, udnColumnCounter];
				END_FOR	
			END_FOR		
			
			udnRowCounter := 0;
			
			etTraceState := ET_TRACE_State_eDataWrite;
		END_IF

	ET_TRACE_State_eGetData:
		IF NOT fbCycleTime.bTimeStarted
		   OR fbCycleTime.stActTime.dwMiliSec >= udnSampleTime * udnWriteCounter
		THEN
			udnRowCounter := GVL_Trace.MAX_TRACE_ROWS;
			udnWriteCounter := udnWriteCounter + 1;
		
			arsValueRecords[udnRowCounter, 0] := UDINT_TO_STRING(udnWriteCounter);
		
			FOR udnColumnCounter := 0 TO GVL_Trace.MAX_TRACE_COLUMNS
			DO 
				IF NOT fbCycleTime.bTimeStarted
				THEN
					fbFileHandler.arsWriteRecords[0, udnColumnCounter] := '';			
				ELSE
					fbFileHandler.arsWriteRecords[0, udnColumnCounter] := arsValueRecords[udnRowCounter, udnColumnCounter];
				END_IF
				
			END_FOR		
			
			etTraceState := ET_TRACE_State_eDataWrite;
		END_IF
	
	ET_TRACE_State_eDataWrite:
		fbFileHandler.bExecute := TRUE;
			
		IF fbFileHandler.bBusy
		   AND NOT fbFileHandler.bError
		THEN
			etTraceState := ET_TRACE_State_eWfDataWrite;
			
		ELSIF fbFileHandler.bError
		THEN
			fbFileHandler.bExecute := FALSE;

			etTraceState := ET_TRACE_State_eError;
		END_IF
		
	ET_TRACE_State_eWfDataWrite:
		IF fbFileHandler.bDone
		    AND NOT fbFileHandler.bError
		THEN
			fbFileHandler.bExecute := FALSE;
		
			IF fbCycleTime.bTimeStarted
			THEN	
				etTraceState := ET_TRACE_State_eGetData;
			ELSE
				etTraceState := ET_TRACE_State_eDone;	
			END_IF
			
		ELSIF fbFileHandler.bError
		THEN
			fbFileHandler.bExecute := FALSE;

			etTraceState := ET_TRACE_State_eError;
		END_IF

	ET_Trace_State_eDone:
		bBusy := FALSE;
		bDone := TRUE;
		bError := FALSE;
		
		etTraceState := ET_TRACE_State_eNoExecute;					(* Next step *)

	ET_Trace_State_eError:
		bBusy := FALSE;
		bDone := FALSE;
		bError := TRUE;

		etTraceState := ET_TRACE_State_eNoExecute;					(* Next step *)

	ET_Trace_State_eNoExecute:
		IF NOT bExecute
		THEN
			bBusy := FALSE;
			bDone := FALSE;
			bError := FALSE;

			etTraceState := ET_TRACE_State_eWaitExecute;			(* Next step *)

		END_IF		
END_CASE

END_FUNCTION_BLOCK

// ---- POUs/Tc3 Objects/Traceability/FB_TraceSingle.TcPOU
FUNCTION_BLOCK FB_TraceSingle
(*

This function block is used to traceability of data.

Constructor: 		Patryk Panylo
Company:		E. Riexinger GmbH
Date:			02.09.2016
Version:			1.00

Date:			Revision:		Who:				Comment
21.02.2018		0.01			PPA						Additional logger for samples

*)
VAR_INPUT
	(* Input variables / Eingang Variablen *)
	bEnable						:BOOL;					(* Enable FB *)
	sFilePath					:STRING := 'C:\Riex\Traceability\NewData\';	(* Path to file e.g. 'c:\', \Hard Disk\ *)
	sFileName					:STRING := 'default';	(* Name of file *)
	bExecute					:BOOL;					(* Execute write data *)
	bReset						:BOOL;					(* Reset write data *)	
	arsNameRecords				:ARRAY[0..GVL_Trace.MAX_TRACE_ROWS, 0..GVL_Trace.MAX_TRACE_COLUMNS] OF STRING(GVL_Trace.MAX_TRACE_FIELD_LENGTH);
	arsValueRecords				:ARRAY[0..GVL_Trace.MAX_TRACE_ROWS, 0..GVL_Trace.MAX_TRACE_COLUMNS] OF STRING(GVL_Trace.MAX_TRACE_FIELD_LENGTH);
	tTimeout					:TIME := T#1S;			(* States the time before the function is cancelled *)
END_VAR
VAR_OUTPUT
	(* Output variables / Ausgang Variablen *)
	bBusy						:BOOL;					(* Program busy *)
	bDone						:BOOL;					(* Program done *)
	bError						:BOOL;					(* Program error *)
	udnErrNo					:UDINT;					(* Error number *)
END_VAR
VAR_IN_OUT
	fbFileHandler				:FB_FileCSVHandler;				(* Traceability *)
END_VAR
VAR
	(* Enummerations *)
	etTraceState				:ET_TRACE_State := ET_TRACE_State_eWaitExecute;
	
	(* Variables *)
	udnWriteCounter				:UDINT;
	
	sLastFilePath				:STRING;
	sLastFileName				:STRING;
	
	udnRowCounter				:UDINT;
	udnColumnCounter			:UDINT;

	bFirstTime					:BOOL;					(* First PLC cycle *)

	(* References *)

	(* Interfaces *)

	(* Instances *)
	rtExecute						:R_TRIG;
END_VAR

IF NOT bEnable				(* Enable FB *)
THEN
	bFirstTime := FALSE;		(* First PLC cycle *)
	bBusy := FALSE;			(* Program busy *)
	bDone := FALSE;			(* Program done *)
	bError := FALSE;			(* Program error *)
	udnErrNo := 0;				(* Error number *)
	RETURN;
END_IF

IF NOT bFirstTime
THEN

	bFirstTime := TRUE;
END_IF

IF bReset
   AND bError
THEN
	bBusy := FALSE;
	bDone := FALSE;
	bError := FALSE;
	
	etTraceState := ET_TRACE_State_eWaitExecute;
END_IF

rtExecute(CLK := bExecute);

CASE etTraceState
OF
	ET_TRACE_State_eWaitExecute:
		IF rtExecute.Q
		   AND NOT fbFileHandler.bBusy
		THEN
			bBusy := TRUE;
			bDone := FALSE;
			bError := FALSE;
			udnErrNo := 0;

			fbFileHandler.bExecute := FALSE;
			fbFileHandler.sFilePath := sFilePath;
			fbFileHandler.sFileName := sFileName; 
			
			udnWriteCounter := 0;
			udnRowCounter := 0;
			udnColumnCounter := 0;
			
			IF (sLastFilePath <> sFilePath)
			   OR (sLastFileName <> sFileName)
			THEN
				FOR udnColumnCounter := 0 TO GVL_Trace.MAX_TRACE_COLUMNS
				DO 
					fbFileHandler.arsWriteRecords[0, udnColumnCounter] := arsNameRecords[0, udnColumnCounter];
				END_FOR

				sLastFilePath := sFilePath;
				sLastFileName := sFileName;
				
				etTraceState := ET_TRACE_State_eDataWrite;
			
			ELSE
				udnWriteCounter := udnWriteCounter + 1;
				
				etTraceState := ET_TRACE_State_eGetData;
			END_IF
								
		END_IF

	ET_TRACE_State_eGetData:
		FOR udnColumnCounter := 0 TO GVL_Trace.MAX_TRACE_COLUMNS
		DO 
			fbFileHandler.arsWriteRecords[udnRowCounter, udnColumnCounter] := arsValueRecords[udnRowCounter, udnColumnCounter];
		END_FOR
		
		etTraceState := ET_TRACE_State_eDataWrite;
			
	ET_TRACE_State_eDataWrite:
		fbFileHandler.bExecute := TRUE;

		IF fbFileHandler.bBusy
		   AND NOT fbFileHandler.bError
		THEN
			etTraceState := ET_TRACE_State_eWfDataWrite;
			
		ELSIF fbFileHandler.bError
		THEN
			fbFileHandler.bExecute := FALSE;

			etTraceState := ET_TRACE_State_eError;
		END_IF
		
	ET_TRACE_State_eWfDataWrite:
		IF fbFileHandler.bDone
		    AND NOT fbFileHandler.bError
		THEN
			fbFileHandler.bExecute := FALSE;

			IF udnWriteCounter <= 0
			THEN
				udnWriteCounter := udnWriteCounter + 1;
				
				etTraceState := ET_TRACE_State_eGetData;
			ELSE
				etTraceState := ET_TRACE_State_eDone;
			END_IF
			
		ELSIF fbFileHandler.bError
		THEN
			fbFileHandler.bExecute := FALSE;

			etTraceState := ET_TRACE_State_eError;
		END_IF

	ET_TRACE_State_eDone:
		bBusy := FALSE;
		bDone := TRUE;
		bError := FALSE;
		
		etTraceState := ET_TRACE_State_eNoExecute;					(* Next step *)

	ET_TRACE_State_eError:
		bBusy := FALSE;
		bDone := FALSE;
		bError := TRUE;

		etTraceState := ET_TRACE_State_eNoExecute;					(* Next step *)

	ET_TRACE_State_eNoExecute:
		IF NOT bExecute
		THEN
			bBusy := FALSE;
			bDone := FALSE;
			bError := FALSE;

			etTraceState := ET_TRACE_State_eWaitExecute;			(* Next step *)

		END_IF		
END_CASE

END_FUNCTION_BLOCK
